(* IEC 61131-3 sources: veristc/veri-stc/tests/st-examples (part 2) *)

cond_a := LimitHigh(raw_030_a, 130);
cond_a := cond_a AND quality_a;
cond_a := cond_a AND (NOT bypass_a);
input_valid_a := InputValid(raw_030_a, 0, 1000);
cond_a := cond_a AND input_valid_a;
IF NOT input_valid_a THEN
    channel_fault_a := channel_fault_a + 1;
END_IF;
cond_b := LimitHigh(raw_030_b, 130);
cond_b := cond_b AND quality_b;
cond_b := cond_b AND (NOT bypass_b);
input_valid_b := InputValid(raw_030_b, 0, 1000);
cond_b := cond_b AND input_valid_b;
IF NOT input_valid_b THEN
    channel_fault_b := channel_fault_b + 1;
END_IF;
cond_c := LimitHigh(raw_030_c, 130);
cond_c := cond_c AND quality_c;
cond_c := cond_c AND (NOT bypass_c);
input_valid_c := InputValid(raw_030_c, 0, 1000);
cond_c := cond_c AND input_valid_c;
IF NOT input_valid_c THEN
    channel_fault_c := channel_fault_c + 1;
END_IF;
cond_d := LimitHigh(raw_030_d, 130);
cond_d := cond_d AND quality_d;
cond_d := cond_d AND (NOT bypass_d);
input_valid_d := InputValid(raw_030_d, 0, 1000);
cond_d := cond_d AND input_valid_d;
IF NOT input_valid_d THEN
    channel_fault_d := channel_fault_d + 1;
END_IF;
vote_ok := TwoOfFour(cond_a, cond_b, cond_c, cond_d);
IF cond_a <> cond_b THEN
    diagnosis_count := diagnosis_count + 1;
END_IF;
IF cond_c <> cond_d THEN
    diagnosis_count := diagnosis_count + 1;
END_IF;
IF NOT vote_ok THEN
    diagnosis_count := diagnosis_count + 1;
END_IF;
latch_a_030 := RS_Next(vote_ok, train_a_reset, latch_a_030);
IF latch_a_030 AND (NOT train_a_inhibit) THEN
    mask_a_03 := mask_a_03 + 64;
    trip_a := 0 < 1;
    scram_a := 0 < 1;
    breaker_a := 0 > 1;
    mfw_a := 0 < 1;
    alarm_a := 0 < 1;
END_IF;
latch_b_030 := RS_Next(vote_ok, train_b_reset, latch_b_030);
IF latch_b_030 AND (NOT train_b_inhibit) THEN
    mask_b_03 := mask_b_03 + 64;
    trip_b := 0 < 1;
    scram_b := 0 < 1;
    breaker_b := 0 > 1;
    mfw_b := 0 < 1;
    alarm_b := 0 < 1;
END_IF;
IF (raw_030_a > 130) AND (NOT cond_a) THEN
    channel_fault_a := channel_fault_a + 1;
END_IF;
IF (raw_030_b > 130) AND (NOT cond_b) THEN
    channel_fault_b := channel_fault_b + 1;
END_IF;
IF (raw_030_c > 130) AND (NOT cond_c) THEN
    channel_fault_c := channel_fault_c + 1;
END_IF;
IF (raw_030_d > 130) AND (NOT cond_d) THEN
    channel_fault_d := channel_fault_d + 1;
END_IF;
IF vote_ok AND train_a_inhibit THEN
    diagnosis_count := diagnosis_count + 1;
END_IF;
IF vote_ok AND train_b_inhibit THEN
    diagnosis_count := diagnosis_count + 1;
END_IF;

cond_a := LimitHigh(raw_031_a, 131);
cond_a := cond_a AND quality_a;
cond_a := cond_a AND (NOT bypass_a);
input_valid_a := InputValid(raw_031_a, 0, 1000);
cond_a := cond_a AND input_valid_a;
IF NOT input_valid_a THEN
    channel_fault_a := channel_fault_a + 1;
END_IF;
cond_b := LimitHigh(raw_031_b, 131);
cond_b := cond_b AND quality_b;
cond_b := cond_b AND (NOT bypass_b);
input_valid_b := InputValid(raw_031_b, 0, 1000);
cond_b := cond_b AND input_valid_b;
IF NOT input_valid_b THEN
    channel_fault_b := channel_fault_b + 1;
END_IF;
cond_c := LimitHigh(raw_031_c, 131);
cond_c := cond_c AND quality_c;
cond_c := cond_c AND (NOT bypass_c);
input_valid_c := InputValid(raw_031_c, 0, 1000);
cond_c := cond_c AND input_valid_c;
IF NOT input_valid_c THEN
    channel_fault_c := channel_fault_c + 1;
END_IF;
cond_d := LimitHigh(raw_031_d, 131);
cond_d := cond_d AND quality_d;
cond_d := cond_d AND (NOT bypass_d);
input_valid_d := InputValid(raw_031_d, 0, 1000);
cond_d := cond_d AND input_valid_d;
IF NOT input_valid_d THEN
    channel_fault_d := channel_fault_d + 1;
END_IF;
vote_ok := TwoOfFour(cond_a, cond_b, cond_c, cond_d);
IF cond_a <> cond_b THEN
    diagnosis_count := diagnosis_count + 1;
END_IF;
IF cond_c <> cond_d THEN
    diagnosis_count := diagnosis_count + 1;
END_IF;
IF NOT vote_ok THEN
    diagnosis_count := diagnosis_count + 1;
END_IF;
latch_a_031 := RS_Next(vote_ok, train_a_reset, latch_a_031);
IF latch_a_031 AND (NOT train_a_inhibit) THEN
    mask_a_03 := mask_a_03 + 128;
    trip_a := 0 < 1;
    scram_a := 0 < 1;
    breaker_a := 0 > 1;
    afw_a := 0 < 1;
    alarm_a := 0 < 1;
END_IF;
latch_b_031 := RS_Next(vote_ok, train_b_reset, latch_b_031);
IF latch_b_031 AND (NOT train_b_inhibit) THEN
    mask_b_03 := mask_b_03 + 128;
    trip_b := 0 < 1;
    scram_b := 0 < 1;
    breaker_b := 0 > 1;
    afw_b := 0 < 1;
    alarm_b := 0 < 1;
END_IF;
IF (raw_031_a > 131) AND (NOT cond_a) THEN
    channel_fault_a := channel_fault_a + 1;
END_IF;
IF (raw_031_b > 131) AND (NOT cond_b) THEN
    channel_fault_b := channel_fault_b + 1;
END_IF;
IF (raw_031_c > 131) AND (NOT cond_c) THEN
    channel_fault_c := channel_fault_c + 1;
END_IF;
IF (raw_031_d > 131) AND (NOT cond_d) THEN
    channel_fault_d := channel_fault_d + 1;
END_IF;
IF vote_ok AND train_a_inhibit THEN
    diagnosis_count := diagnosis_count + 1;
END_IF;
IF vote_ok AND train_b_inhibit THEN
    diagnosis_count := diagnosis_count + 1;
END_IF;

cond_a := LimitHigh(raw_032_a, 132);
cond_a := cond_a AND quality_a;
cond_a := cond_a AND (NOT bypass_a);
input_valid_a := InputValid(raw_032_a, 0, 1000);
cond_a := cond_a AND input_valid_a;
IF NOT input_valid_a THEN
    channel_fault_a := channel_fault_a + 1;
END_IF;
cond_b := LimitHigh(raw_032_b, 132);
cond_b := cond_b AND quality_b;
cond_b := cond_b AND (NOT bypass_b);
input_valid_b := InputValid(raw_032_b, 0, 1000);
cond_b := cond_b AND input_valid_b;
IF NOT input_valid_b THEN
    channel_fault_b := channel_fault_b + 1;
END_IF;
cond_c := LimitHigh(raw_032_c, 132);
cond_c := cond_c AND quality_c;
cond_c := cond_c AND (NOT bypass_c);
input_valid_c := InputValid(raw_032_c, 0, 1000);
cond_c := cond_c AND input_valid_c;
IF NOT input_valid_c THEN
    channel_fault_c := channel_fault_c + 1;
END_IF;
cond_d := LimitHigh(raw_032_d, 132);
cond_d := cond_d AND quality_d;
cond_d := cond_d AND (NOT bypass_d);
input_valid_d := InputValid(raw_032_d, 0, 1000);
cond_d := cond_d AND input_valid_d;
IF NOT input_valid_d THEN
    channel_fault_d := channel_fault_d + 1;
END_IF;
vote_ok := TwoOfFour(cond_a, cond_b, cond_c, cond_d);
IF cond_a <> cond_b THEN
    diagnosis_count := diagnosis_count + 1;
END_IF;
IF cond_c <> cond_d THEN
    diagnosis_count := diagnosis_count + 1;
END_IF;
IF NOT vote_ok THEN
    diagnosis_count := diagnosis_count + 1;
END_IF;
latch_a_032 := RS_Next(vote_ok, train_a_reset, latch_a_032);
IF latch_a_032 AND (NOT train_a_inhibit) THEN
    mask_a_04 := mask_a_04 + 1;
    trip_a := 0 < 1;
    scram_a := 0 < 1;
    breaker_a := 0 > 1;
    si_a := 0 < 1;
    alarm_a := 0 < 1;
END_IF;
latch_b_032 := RS_Next(vote_ok, train_b_reset, latch_b_032);
IF latch_b_032 AND (NOT train_b_inhibit) THEN
    mask_b_04 := mask_b_04 + 1;
    trip_b := 0 < 1;
    scram_b := 0 < 1;
    breaker_b := 0 > 1;
    si_b := 0 < 1;
    alarm_b := 0 < 1;
END_IF;
IF (raw_032_a > 132) AND (NOT cond_a) THEN
    channel_fault_a := channel_fault_a + 1;
END_IF;
IF (raw_032_b > 132) AND (NOT cond_b) THEN
    channel_fault_b := channel_fault_b + 1;
END_IF;
IF (raw_032_c > 132) AND (NOT cond_c) THEN
    channel_fault_c := channel_fault_c + 1;
END_IF;
IF (raw_032_d > 132) AND (NOT cond_d) THEN
    channel_fault_d := channel_fault_d + 1;
END_IF;
IF vote_ok AND train_a_inhibit THEN
    diagnosis_count := diagnosis_count + 1;
END_IF;
IF vote_ok AND train_b_inhibit THEN
    diagnosis_count := diagnosis_count + 1;
END_IF;

cond_a := LimitHigh(raw_033_a, 133);
cond_a := cond_a AND quality_a;
cond_a := cond_a AND (NOT bypass_a);
input_valid_a := InputValid(raw_033_a, 0, 1000);
cond_a := cond_a AND input_valid_a;
IF NOT input_valid_a THEN
    channel_fault_a := channel_fault_a + 1;
END_IF;
cond_b := LimitHigh(raw_033_b, 133);
cond_b := cond_b AND quality_b;
cond_b := cond_b AND (NOT bypass_b);
input_valid_b := InputValid(raw_033_b, 0, 1000);
cond_b := cond_b AND input_valid_b;
IF NOT input_valid_b THEN
    channel_fault_b := channel_fault_b + 1;
END_IF;
cond_c := LimitHigh(raw_033_c, 133);
cond_c := cond_c AND quality_c;
cond_c := cond_c AND (NOT bypass_c);
input_valid_c := InputValid(raw_033_c, 0, 1000);
cond_c := cond_c AND input_valid_c;
IF NOT input_valid_c THEN
    channel_fault_c := channel_fault_c + 1;
END_IF;
cond_d := LimitHigh(raw_033_d, 133);
cond_d := cond_d AND quality_d;
cond_d := cond_d AND (NOT bypass_d);
input_valid_d := InputValid(raw_033_d, 0, 1000);
cond_d := cond_d AND input_valid_d;
IF NOT input_valid_d THEN
    channel_fault_d := channel_fault_d + 1;
END_IF;
vote_ok := TwoOfFour(cond_a, cond_b, cond_c, cond_d);
IF cond_a <> cond_b THEN
    diagnosis_count := diagnosis_count + 1;
END_IF;
IF cond_c <> cond_d THEN
    diagnosis_count := diagnosis_count + 1;
END_IF;
IF NOT vote_ok THEN
    diagnosis_count := diagnosis_count + 1;
END_IF;
latch_a_033 := RS_Next(vote_ok, train_a_reset, latch_a_033);
IF latch_a_033 AND (NOT train_a_inhibit) THEN
    mask_a_04 := mask_a_04 + 2;
    trip_a := 0 < 1;
    scram_a := 0 < 1;
    breaker_a := 0 > 1;
    ci_a := 0 < 1;
    alarm_a := 0 < 1;
END_IF;
latch_b_033 := RS_Next(vote_ok, train_b_reset, latch_b_033);
IF latch_b_033 AND (NOT train_b_inhibit) THEN
    mask_b_04 := mask_b_04 + 2;
    trip_b := 0 < 1;
    scram_b := 0 < 1;
    breaker_b := 0 > 1;
    ci_b := 0 < 1;
    alarm_b := 0 < 1;
END_IF;
IF (raw_033_a > 133) AND (NOT cond_a) THEN
    channel_fault_a := channel_fault_a + 1;
END_IF;
IF (raw_033_b > 133) AND (NOT cond_b) THEN
    channel_fault_b := channel_fault_b + 1;
END_IF;
IF (raw_033_c > 133) AND (NOT cond_c) THEN
    channel_fault_c := channel_fault_c + 1;
END_IF;
IF (raw_033_d > 133) AND (NOT cond_d) THEN
    channel_fault_d := channel_fault_d + 1;
END_IF;
IF vote_ok AND train_a_inhibit THEN
    diagnosis_count := diagnosis_count + 1;
END_IF;
IF vote_ok AND train_b_inhibit THEN
    diagnosis_count := diagnosis_count + 1;
END_IF;

cond_a := LimitHigh(raw_034_a, 134);
cond_a := cond_a AND quality_a;
cond_a := cond_a AND (NOT bypass_a);
input_valid_a := InputValid(raw_034_a, 0, 1000);
cond_a := cond_a AND input_valid_a;
IF NOT input_valid_a THEN
    channel_fault_a := channel_fault_a + 1;
END_IF;
cond_b := LimitHigh(raw_034_b, 134);
cond_b := cond_b AND quality_b;
cond_b := cond_b AND (NOT bypass_b);
input_valid_b := InputValid(raw_034_b, 0, 1000);
cond_b := cond_b AND input_valid_b;
IF NOT input_valid_b THEN
    channel_fault_b := channel_fault_b + 1;
END_IF;
cond_c := LimitHigh(raw_034_c, 134);
cond_c := cond_c AND quality_c;
cond_c := cond_c AND (NOT bypass_c);
input_valid_c := InputValid(raw_034_c, 0, 1000);
cond_c := cond_c AND input_valid_c;
IF NOT input_valid_c THEN
    channel_fault_c := channel_fault_c + 1;
END_IF;
cond_d := LimitHigh(raw_034_d, 134);
cond_d := cond_d AND quality_d;
cond_d := cond_d AND (NOT bypass_d);
input_valid_d := InputValid(raw_034_d, 0, 1000);
cond_d := cond_d AND input_valid_d;
IF NOT input_valid_d THEN
    channel_fault_d := channel_fault_d + 1;
END_IF;
vote_ok := TwoOfFour(cond_a, cond_b, cond_c, cond_d);
IF cond_a <> cond_b THEN
    diagnosis_count := diagnosis_count + 1;
END_IF;
IF cond_c <> cond_d THEN
    diagnosis_count := diagnosis_count + 1;
END_IF;
IF NOT vote_ok THEN
    diagnosis_count := diagnosis_count + 1;
END_IF;
latch_a_034 := RS_Next(vote_ok, train_a_reset, latch_a_034);
IF latch_a_034 AND (NOT train_a_inhibit) THEN
    mask_a_04 := mask_a_04 + 4;
    trip_a := 0 < 1;
    scram_a := 0 < 1;
    breaker_a := 0 > 1;
    mfw_a := 0 < 1;
    alarm_a := 0 < 1;
END_IF;
latch_b_034 := RS_Next(vote_ok, train_b_reset, latch_b_034);
IF latch_b_034 AND (NOT train_b_inhibit) THEN
    mask_b_04 := mask_b_04 + 4;
    trip_b := 0 < 1;
    scram_b := 0 < 1;
    breaker_b := 0 > 1;
    mfw_b := 0 < 1;
    alarm_b := 0 < 1;
END_IF;
IF (raw_034_a > 134) AND (NOT cond_a) THEN
    channel_fault_a := channel_fault_a + 1;
END_IF;
IF (raw_034_b > 134) AND (NOT cond_b) THEN
    channel_fault_b := channel_fault_b + 1;
END_IF;
IF (raw_034_c > 134) AND (NOT cond_c) THEN
    channel_fault_c := channel_fault_c + 1;
END_IF;
IF (raw_034_d > 134) AND (NOT cond_d) THEN
    channel_fault_d := channel_fault_d + 1;
END_IF;
IF vote_ok AND train_a_inhibit THEN
    diagnosis_count := diagnosis_count + 1;
END_IF;
IF vote_ok AND train_b_inhibit THEN
    diagnosis_count := diagnosis_count + 1;
END_IF;

cond_a := LimitHigh(raw_035_a, 135);
cond_a := cond_a AND quality_a;
cond_a := cond_a AND (NOT bypass_a);
input_valid_a := InputValid(raw_035_a, 0, 1000);
cond_a := cond_a AND input_valid_a;
IF NOT input_valid_a THEN
    channel_fault_a := channel_fault_a + 1;
END_IF;
cond_b := LimitHigh(raw_035_b, 135);
cond_b := cond_b AND quality_b;
cond_b := cond_b AND (NOT bypass_b);
input_valid_b := InputValid(raw_035_b, 0, 1000);
cond_b := cond_b AND input_valid_b;
IF NOT input_valid_b THEN
    channel_fault_b := channel_fault_b + 1;
END_IF;
cond_c := LimitHigh(raw_035_c, 135);
cond_c := cond_c AND quality_c;
cond_c := cond_c AND (NOT bypass_c);
input_valid_c := InputValid(raw_035_c, 0, 1000);
cond_c := cond_c AND input_valid_c;
IF NOT input_valid_c THEN
    channel_fault_c := channel_fault_c + 1;
END_IF;
cond_d := LimitHigh(raw_035_d, 135);
cond_d := cond_d AND quality_d;
cond_d := cond_d AND (NOT bypass_d);
input_valid_d := InputValid(raw_035_d, 0, 1000);
cond_d := cond_d AND input_valid_d;
IF NOT input_valid_d THEN
    channel_fault_d := channel_fault_d + 1;
END_IF;
vote_ok := TwoOfFour(cond_a, cond_b, cond_c, cond_d);
IF cond_a <> cond_b THEN
    diagnosis_count := diagnosis_count + 1;
END_IF;
IF cond_c <> cond_d THEN
    diagnosis_count := diagnosis_count + 1;
END_IF;
IF NOT vote_ok THEN
    diagnosis_count := diagnosis_count + 1;
END_IF;
latch_a_035 := RS_Next(vote_ok, train_a_reset, latch_a_035);
IF latch_a_035 AND (NOT train_a_inhibit) THEN
    mask_a_04 := mask_a_04 + 8;
    trip_a := 0 < 1;
    scram_a := 0 < 1;
    breaker_a := 0 > 1;
    afw_a := 0 < 1;
    alarm_a := 0 < 1;
END_IF;
latch_b_035 := RS_Next(vote_ok, train_b_reset, latch_b_035);
IF latch_b_035 AND (NOT train_b_inhibit) THEN
    mask_b_04 := mask_b_04 + 8;
    trip_b := 0 < 1;
    scram_b := 0 < 1;
    breaker_b := 0 > 1;
    afw_b := 0 < 1;
    alarm_b := 0 < 1;
END_IF;
IF (raw_035_a > 135) AND (NOT cond_a) THEN
    channel_fault_a := channel_fault_a + 1;
END_IF;
IF (raw_035_b > 135) AND (NOT cond_b) THEN
    channel_fault_b := channel_fault_b + 1;
END_IF;
IF (raw_035_c > 135) AND (NOT cond_c) THEN
    channel_fault_c := channel_fault_c + 1;
END_IF;
IF (raw_035_d > 135) AND (NOT cond_d) THEN
    channel_fault_d := channel_fault_d + 1;
END_IF;
IF vote_ok AND train_a_inhibit THEN
    diagnosis_count := diagnosis_count + 1;
END_IF;
IF vote_ok AND train_b_inhibit THEN
    diagnosis_count := diagnosis_count + 1;
END_IF;

cond_a := LimitHigh(raw_036_a, 136);
cond_a := cond_a AND quality_a;
cond_a := cond_a AND (NOT bypass_a);
input_valid_a := InputValid(raw_036_a, 0, 1000);
cond_a := cond_a AND input_valid_a;
IF NOT input_valid_a THEN
    channel_fault_a := channel_fault_a + 1;
END_IF;
cond_b := LimitHigh(raw_036_b, 136);
cond_b := cond_b AND quality_b;
cond_b := cond_b AND (NOT bypass_b);
input_valid_b := InputValid(raw_036_b, 0, 1000);
cond_b := cond_b AND input_valid_b;
IF NOT input_valid_b THEN
    channel_fault_b := channel_fault_b + 1;
END_IF;
cond_c := LimitHigh(raw_036_c, 136);
cond_c := cond_c AND quality_c;
cond_c := cond_c AND (NOT bypass_c);
input_valid_c := InputValid(raw_036_c, 0, 1000);
cond_c := cond_c AND input_valid_c;
IF NOT input_valid_c THEN
    channel_fault_c := channel_fault_c + 1;
END_IF;
cond_d := LimitHigh(raw_036_d, 136);
cond_d := cond_d AND quality_d;
cond_d := cond_d AND (NOT bypass_d);
input_valid_d := InputValid(raw_036_d, 0, 1000);
cond_d := cond_d AND input_valid_d;
IF NOT input_valid_d THEN
    channel_fault_d := channel_fault_d + 1;
END_IF;
vote_ok := TwoOfFour(cond_a, cond_b, cond_c, cond_d);
IF cond_a <> cond_b THEN
    diagnosis_count := diagnosis_count + 1;
END_IF;
IF cond_c <> cond_d THEN
    diagnosis_count := diagnosis_count + 1;
END_IF;
IF NOT vote_ok THEN
    diagnosis_count := diagnosis_count + 1;
END_IF;
latch_a_036 := RS_Next(vote_ok, train_a_reset, latch_a_036);
IF latch_a_036 AND (NOT train_a_inhibit) THEN
    mask_a_04 := mask_a_04 + 16;
    trip_a := 0 < 1;
    scram_a := 0 < 1;
    breaker_a := 0 > 1;
    si_a := 0 < 1;
    alarm_a := 0 < 1;
END_IF;
latch_b_036 := RS_Next(vote_ok, train_b_reset, latch_b_036);
IF latch_b_036 AND (NOT train_b_inhibit) THEN
    mask_b_04 := mask_b_04 + 16;
    trip_b := 0 < 1;
    scram_b := 0 < 1;
    breaker_b := 0 > 1;
    si_b := 0 < 1;
    alarm_b := 0 < 1;
END_IF;
IF (raw_036_a > 136) AND (NOT cond_a) THEN
    channel_fault_a := channel_fault_a + 1;
END_IF;
IF (raw_036_b > 136) AND (NOT cond_b) THEN
    channel_fault_b := channel_fault_b + 1;
END_IF;
IF (raw_036_c > 136) AND (NOT cond_c) THEN
    channel_fault_c := channel_fault_c + 1;
END_IF;
IF (raw_036_d > 136) AND (NOT cond_d) THEN
    channel_fault_d := channel_fault_d + 1;
END_IF;
IF vote_ok AND train_a_inhibit THEN
    diagnosis_count := diagnosis_count + 1;
END_IF;
IF vote_ok AND train_b_inhibit THEN
    diagnosis_count := diagnosis_count + 1;
END_IF;

cond_a := LimitHigh(raw_037_a, 137);
cond_a := cond_a AND quality_a;
cond_a := cond_a AND (NOT bypass_a);
input_valid_a := InputValid(raw_037_a, 0, 1000);
cond_a := cond_a AND input_valid_a;
IF NOT input_valid_a THEN
    channel_fault_a := channel_fault_a + 1;
END_IF;
cond_b := LimitHigh(raw_037_b, 137);
cond_b := cond_b AND quality_b;
cond_b := cond_b AND (NOT bypass_b);
input_valid_b := InputValid(raw_037_b, 0, 1000);
cond_b := cond_b AND input_valid_b;
IF NOT input_valid_b THEN
    channel_fault_b := channel_fault_b + 1;
END_IF;
cond_c := LimitHigh(raw_037_c, 137);
cond_c := cond_c AND quality_c;
cond_c := cond_c AND (NOT bypass_c);
input_valid_c := InputValid(raw_037_c, 0, 1000);
cond_c := cond_c AND input_valid_c;
IF NOT input_valid_c THEN
    channel_fault_c := channel_fault_c + 1;
END_IF;
cond_d := LimitHigh(raw_037_d, 137);
cond_d := cond_d AND quality_d;
cond_d := cond_d AND (NOT bypass_d);
input_valid_d := InputValid(raw_037_d, 0, 1000);
cond_d := cond_d AND input_valid_d;
IF NOT input_valid_d THEN
    channel_fault_d := channel_fault_d + 1;
END_IF;
vote_ok := TwoOfFour(cond_a, cond_b, cond_c, cond_d);
IF cond_a <> cond_b THEN
    diagnosis_count := diagnosis_count + 1;
END_IF;
IF cond_c <> cond_d THEN
    diagnosis_count := diagnosis_count + 1;
END_IF;
IF NOT vote_ok THEN
    diagnosis_count := diagnosis_count + 1;
END_IF;
latch_a_037 := RS_Next(vote_ok, train_a_reset, latch_a_037);
IF latch_a_037 AND (NOT train_a_inhibit) THEN
    mask_a_04 := mask_a_04 + 32;
    trip_a := 0 < 1;
    scram_a := 0 < 1;
    breaker_a := 0 > 1;
    ci_a := 0 < 1;
    alarm_a := 0 < 1;
END_IF;
latch_b_037 := RS_Next(vote_ok, train_b_reset, latch_b_037);
IF latch_b_037 AND (NOT train_b_inhibit) THEN
    mask_b_04 := mask_b_04 + 32;
    trip_b := 0 < 1;
    scram_b := 0 < 1;
    breaker_b := 0 > 1;
    ci_b := 0 < 1;
    alarm_b := 0 < 1;
END_IF;
IF (raw_037_a > 137) AND (NOT cond_a) THEN
    channel_fault_a := channel_fault_a + 1;
END_IF;
IF (raw_037_b > 137) AND (NOT cond_b) THEN
    channel_fault_b := channel_fault_b + 1;
END_IF;
IF (raw_037_c > 137) AND (NOT cond_c) THEN
    channel_fault_c := channel_fault_c + 1;
END_IF;
IF (raw_037_d > 137) AND (NOT cond_d) THEN
    channel_fault_d := channel_fault_d + 1;
END_IF;
IF vote_ok AND train_a_inhibit THEN
    diagnosis_count := diagnosis_count + 1;
END_IF;
IF vote_ok AND train_b_inhibit THEN
    diagnosis_count := diagnosis_count + 1;
END_IF;

cond_a := LimitHigh(raw_038_a, 138);
cond_a := cond_a AND quality_a;
cond_a := cond_a AND (NOT bypass_a);
input_valid_a := InputValid(raw_038_a, 0, 1000);
cond_a := cond_a AND input_valid_a;
IF NOT input_valid_a THEN
    channel_fault_a := channel_fault_a + 1;
END_IF;
cond_b := LimitHigh(raw_038_b, 138);
cond_b := cond_b AND quality_b;
cond_b := cond_b AND (NOT bypass_b);
input_valid_b := InputValid(raw_038_b, 0, 1000);
cond_b := cond_b AND input_valid_b;
IF NOT input_valid_b THEN
    channel_fault_b := channel_fault_b + 1;
END_IF;
cond_c := LimitHigh(raw_038_c, 138);
cond_c := cond_c AND quality_c;
cond_c := cond_c AND (NOT bypass_c);
input_valid_c := InputValid(raw_038_c, 0, 1000);
cond_c := cond_c AND input_valid_c;
IF NOT input_valid_c THEN
    channel_fault_c := channel_fault_c + 1;
END_IF;
cond_d := LimitHigh(raw_038_d, 138);
cond_d := cond_d AND quality_d;
cond_d := cond_d AND (NOT bypass_d);
input_valid_d := InputValid(raw_038_d, 0, 1000);
cond_d := cond_d AND input_valid_d;
IF NOT input_valid_d THEN
    channel_fault_d := channel_fault_d + 1;
END_IF;
vote_ok := TwoOfFour(cond_a, cond_b, cond_c, cond_d);
IF cond_a <> cond_b THEN
    diagnosis_count := diagnosis_count + 1;
END_IF;
IF cond_c <> cond_d THEN
    diagnosis_count := diagnosis_count + 1;
END_IF;
IF NOT vote_ok THEN
    diagnosis_count := diagnosis_count + 1;
END_IF;
latch_a_038 := RS_Next(vote_ok, train_a_reset, latch_a_038);
IF latch_a_038 AND (NOT train_a_inhibit) THEN
    mask_a_04 := mask_a_04 + 64;
    trip_a := 0 < 1;
    scram_a := 0 < 1;
    breaker_a := 0 > 1;
    mfw_a := 0 < 1;
    alarm_a := 0 < 1;
END_IF;
latch_b_038 := RS_Next(vote_ok, train_b_reset, latch_b_038);
IF latch_b_038 AND (NOT train_b_inhibit) THEN
    mask_b_04 := mask_b_04 + 64;
    trip_b := 0 < 1;
    scram_b := 0 < 1;
    breaker_b := 0 > 1;
    mfw_b := 0 < 1;
    alarm_b := 0 < 1;
END_IF;
IF (raw_038_a > 138) AND (NOT cond_a) THEN
    channel_fault_a := channel_fault_a + 1;
END_IF;
IF (raw_038_b > 138) AND (NOT cond_b) THEN
    channel_fault_b := channel_fault_b + 1;
END_IF;
IF (raw_038_c > 138) AND (NOT cond_c) THEN
    channel_fault_c := channel_fault_c + 1;
END_IF;
IF (raw_038_d > 138) AND (NOT cond_d) THEN
    channel_fault_d := channel_fault_d + 1;
END_IF;
IF vote_ok AND train_a_inhibit THEN
    diagnosis_count := diagnosis_count + 1;
END_IF;
IF vote_ok AND train_b_inhibit THEN
    diagnosis_count := diagnosis_count + 1;
END_IF;

cond_a := LimitHigh(raw_039_a, 139);
cond_a := cond_a AND quality_a;
cond_a := cond_a AND (NOT bypass_a);
input_valid_a := InputValid(raw_039_a, 0, 1000);
cond_a := cond_a AND input_valid_a;
IF NOT input_valid_a THEN
    channel_fault_a := channel_fault_a + 1;
END_IF;
cond_b := LimitHigh(raw_039_b, 139);
cond_b := cond_b AND quality_b;
cond_b := cond_b AND (NOT bypass_b);
input_valid_b := InputValid(raw_039_b, 0, 1000);
cond_b := cond_b AND input_valid_b;
IF NOT input_valid_b THEN
    channel_fault_b := channel_fault_b + 1;
END_IF;
cond_c := LimitHigh(raw_039_c, 139);
cond_c := cond_c AND quality_c;
cond_c := cond_c AND (NOT bypass_c);
input_valid_c := InputValid(raw_039_c, 0, 1000);
cond_c := cond_c AND input_valid_c;
IF NOT input_valid_c THEN
    channel_fault_c := channel_fault_c + 1;
END_IF;
cond_d := LimitHigh(raw_039_d, 139);
cond_d := cond_d AND quality_d;
cond_d := cond_d AND (NOT bypass_d);
input_valid_d := InputValid(raw_039_d, 0, 1000);
cond_d := cond_d AND input_valid_d;
IF NOT input_valid_d THEN
    channel_fault_d := channel_fault_d + 1;
END_IF;
vote_ok := TwoOfFour(cond_a, cond_b, cond_c, cond_d);
IF cond_a <> cond_b THEN
    diagnosis_count := diagnosis_count + 1;
END_IF;
IF cond_c <> cond_d THEN
    diagnosis_count := diagnosis_count + 1;
END_IF;
IF NOT vote_ok THEN
    diagnosis_count := diagnosis_count + 1;
END_IF;
latch_a_039 := RS_Next(vote_ok, train_a_reset, latch_a_039);
IF latch_a_039 AND (NOT train_a_inhibit) THEN
    mask_a_04 := mask_a_04 + 128;
    trip_a := 0 < 1;
    scram_a := 0 < 1;
    breaker_a := 0 > 1;
    afw_a := 0 < 1;
    alarm_a := 0 < 1;
END_IF;
latch_b_039 := RS_Next(vote_ok, train_b_reset, latch_b_039);
IF latch_b_039 AND (NOT train_b_inhibit) THEN
    mask_b_04 := mask_b_04 + 128;
    trip_b := 0 < 1;
    scram_b := 0 < 1;
    breaker_b := 0 > 1;
    afw_b := 0 < 1;
    alarm_b := 0 < 1;
END_IF;
IF (raw_039_a > 139) AND (NOT cond_a) THEN
    channel_fault_a := channel_fault_a + 1;
END_IF;
IF (raw_039_b > 139) AND (NOT cond_b) THEN
    channel_fault_b := channel_fault_b + 1;
END_IF;
IF (raw_039_c > 139) AND (NOT cond_c) THEN
    channel_fault_c := channel_fault_c + 1;
END_IF;
IF (raw_039_d > 139) AND (NOT cond_d) THEN
    channel_fault_d := channel_fault_d + 1;
END_IF;
IF vote_ok AND train_a_inhibit THEN
    diagnosis_count := diagnosis_count + 1;
END_IF;
IF vote_ok AND train_b_inhibit THEN
    diagnosis_count := diagnosis_count + 1;
END_IF;

cond_a := LimitHigh(raw_040_a, 100);
cond_a := cond_a AND quality_a;
cond_a := cond_a AND (NOT bypass_a);
input_valid_a := InputValid(raw_040_a, 0, 1000);
cond_a := cond_a AND input_valid_a;
IF NOT input_valid_a THEN
    channel_fault_a := channel_fault_a + 1;
END_IF;
cond_b := LimitHigh(raw_040_b, 100);
cond_b := cond_b AND quality_b;
cond_b := cond_b AND (NOT bypass_b);
input_valid_b := InputValid(raw_040_b, 0, 1000);
cond_b := cond_b AND input_valid_b;
IF NOT input_valid_b THEN
    channel_fault_b := channel_fault_b + 1;
END_IF;
cond_c := LimitHigh(raw_040_c, 100);
cond_c := cond_c AND quality_c;
cond_c := cond_c AND (NOT bypass_c);
input_valid_c := InputValid(raw_040_c, 0, 1000);
cond_c := cond_c AND input_valid_c;
IF NOT input_valid_c THEN
    channel_fault_c := channel_fault_c + 1;
END_IF;
cond_d := LimitHigh(raw_040_d, 100);
cond_d := cond_d AND quality_d;
cond_d := cond_d AND (NOT bypass_d);
input_valid_d := InputValid(raw_040_d, 0, 1000);
cond_d := cond_d AND input_valid_d;
IF NOT input_valid_d THEN
    channel_fault_d := channel_fault_d + 1;
END_IF;
vote_ok := TwoOfFour(cond_a, cond_b, cond_c, cond_d);
IF cond_a <> cond_b THEN
    diagnosis_count := diagnosis_count + 1;
END_IF;
IF cond_c <> cond_d THEN
    diagnosis_count := diagnosis_count + 1;
END_IF;
IF NOT vote_ok THEN
    diagnosis_count := diagnosis_count + 1;
END_IF;
latch_a_040 := RS_Next(vote_ok, train_a_reset, latch_a_040);
IF latch_a_040 AND (NOT train_a_inhibit) THEN
    mask_a_05 := mask_a_05 + 1;
    trip_a := 0 < 1;
    scram_a := 0 < 1;
    breaker_a := 0 > 1;
    si_a := 0 < 1;
    alarm_a := 0 < 1;
END_IF;
latch_b_040 := RS_Next(vote_ok, train_b_reset, latch_b_040);
IF latch_b_040 AND (NOT train_b_inhibit) THEN
    mask_b_05 := mask_b_05 + 1;
    trip_b := 0 < 1;
    scram_b := 0 < 1;
    breaker_b := 0 > 1;
    si_b := 0 < 1;
    alarm_b := 0 < 1;
END_IF;
IF (raw_040_a > 100) AND (NOT cond_a) THEN
    channel_fault_a := channel_fault_a + 1;
END_IF;
IF (raw_040_b > 100) AND (NOT cond_b) THEN
    channel_fault_b := channel_fault_b + 1;
END_IF;
IF (raw_040_c > 100) AND (NOT cond_c) THEN
    channel_fault_c := channel_fault_c + 1;
END_IF;
IF (raw_040_d > 100) AND (NOT cond_d) THEN
    channel_fault_d := channel_fault_d + 1;
END_IF;
IF vote_ok AND train_a_inhibit THEN
    diagnosis_count := diagnosis_count + 1;
END_IF;
IF vote_ok AND train_b_inhibit THEN
    diagnosis_count := diagnosis_count + 1;
END_IF;

cond_a := LimitHigh(raw_041_a, 101);
cond_a := cond_a AND quality_a;
cond_a := cond_a AND (NOT bypass_a);
input_valid_a := InputValid(raw_041_a, 0, 1000);
cond_a := cond_a AND input_valid_a;
IF NOT input_valid_a THEN
    channel_fault_a := channel_fault_a + 1;
END_IF;
cond_b := LimitHigh(raw_041_b, 101);
cond_b := cond_b AND quality_b;
cond_b := cond_b AND (NOT bypass_b);
input_valid_b := InputValid(raw_041_b, 0, 1000);
cond_b := cond_b AND input_valid_b;
IF NOT input_valid_b THEN
    channel_fault_b := channel_fault_b + 1;
END_IF;
cond_c := LimitHigh(raw_041_c, 101);
cond_c := cond_c AND quality_c;
cond_c := cond_c AND (NOT bypass_c);
input_valid_c := InputValid(raw_041_c, 0, 1000);
cond_c := cond_c AND input_valid_c;
IF NOT input_valid_c THEN
    channel_fault_c := channel_fault_c + 1;
END_IF;
cond_d := LimitHigh(raw_041_d, 101);
cond_d := cond_d AND quality_d;
cond_d := cond_d AND (NOT bypass_d);
input_valid_d := InputValid(raw_041_d, 0, 1000);
cond_d := cond_d AND input_valid_d;
IF NOT input_valid_d THEN
    channel_fault_d := channel_fault_d + 1;
END_IF;
vote_ok := TwoOfFour(cond_a, cond_b, cond_c, cond_d);
IF cond_a <> cond_b THEN
    diagnosis_count := diagnosis_count + 1;
END_IF;
IF cond_c <> cond_d THEN
    diagnosis_count := diagnosis_count + 1;
END_IF;
IF NOT vote_ok THEN
    diagnosis_count := diagnosis_count + 1;
END_IF;
latch_a_041 := RS_Next(vote_ok, train_a_reset, latch_a_041);
IF latch_a_041 AND (NOT train_a_inhibit) THEN
    mask_a_05 := mask_a_05 + 2;
    trip_a := 0 < 1;
    scram_a := 0 < 1;
    breaker_a := 0 > 1;
    ci_a := 0 < 1;
    alarm_a := 0 < 1;
END_IF;
latch_b_041 := RS_Next(vote_ok, train_b_reset, latch_b_041);
IF latch_b_041 AND (NOT train_b_inhibit) THEN
    mask_b_05 := mask_b_05 + 2;
    trip_b := 0 < 1;
    scram_b := 0 < 1;
    breaker_b := 0 > 1;
    ci_b := 0 < 1;
    alarm_b := 0 < 1;
END_IF;
IF (raw_041_a > 101) AND (NOT cond_a) THEN
    channel_fault_a := channel_fault_a + 1;
END_IF;
IF (raw_041_b > 101) AND (NOT cond_b) THEN
    channel_fault_b := channel_fault_b + 1;
END_IF;
IF (raw_041_c > 101) AND (NOT cond_c) THEN
    channel_fault_c := channel_fault_c + 1;
END_IF;
IF (raw_041_d > 101) AND (NOT cond_d) THEN
    channel_fault_d := channel_fault_d + 1;
END_IF;
IF vote_ok AND train_a_inhibit THEN
    diagnosis_count := diagnosis_count + 1;
END_IF;
IF vote_ok AND train_b_inhibit THEN
    diagnosis_count := diagnosis_count + 1;
END_IF;

cond_a := LimitHigh(raw_042_a, 102);
cond_a := cond_a AND quality_a;
cond_a := cond_a AND (NOT bypass_a);
input_valid_a := InputValid(raw_042_a, 0, 1000);
cond_a := cond_a AND input_valid_a;
IF NOT input_valid_a THEN
    channel_fault_a := channel_fault_a + 1;
END_IF;
cond_b := LimitHigh(raw_042_b, 102);
cond_b := cond_b AND quality_b;
cond_b := cond_b AND (NOT bypass_b);
input_valid_b := InputValid(raw_042_b, 0, 1000);
cond_b := cond_b AND input_valid_b;
IF NOT input_valid_b THEN
    channel_fault_b := channel_fault_b + 1;
END_IF;
cond_c := LimitHigh(raw_042_c, 102);
cond_c := cond_c AND quality_c;
cond_c := cond_c AND (NOT bypass_c);
input_valid_c := InputValid(raw_042_c, 0, 1000);
cond_c := cond_c AND input_valid_c;
IF NOT input_valid_c THEN
    channel_fault_c := channel_fault_c + 1;
END_IF;
cond_d := LimitHigh(raw_042_d, 102);
cond_d := cond_d AND quality_d;
cond_d := cond_d AND (NOT bypass_d);
input_valid_d := InputValid(raw_042_d, 0, 1000);
cond_d := cond_d AND input_valid_d;
IF NOT input_valid_d THEN
    channel_fault_d := channel_fault_d + 1;
END_IF;
vote_ok := TwoOfFour(cond_a, cond_b, cond_c, cond_d);
IF cond_a <> cond_b THEN
    diagnosis_count := diagnosis_count + 1;
END_IF;
IF cond_c <> cond_d THEN
    diagnosis_count := diagnosis_count + 1;
END_IF;
IF NOT vote_ok THEN
    diagnosis_count := diagnosis_count + 1;
END_IF;
latch_a_042 := RS_Next(vote_ok, train_a_reset, latch_a_042);
IF latch_a_042 AND (NOT train_a_inhibit) THEN
    mask_a_05 := mask_a_05 + 4;
    trip_a := 0 < 1;
    scram_a := 0 < 1;
    breaker_a := 0 > 1;
    mfw_a := 0 < 1;
    alarm_a := 0 < 1;
END_IF;
latch_b_042 := RS_Next(vote_ok, train_b_reset, latch_b_042);
IF latch_b_042 AND (NOT train_b_inhibit) THEN
    mask_b_05 := mask_b_05 + 4;
    trip_b := 0 < 1;
    scram_b := 0 < 1;
    breaker_b := 0 > 1;
    mfw_b := 0 < 1;
    alarm_b := 0 < 1;
END_IF;
IF (raw_042_a > 102) AND (NOT cond_a) THEN
    channel_fault_a := channel_fault_a + 1;
END_IF;
IF (raw_042_b > 102) AND (NOT cond_b) THEN
    channel_fault_b := channel_fault_b + 1;
END_IF;
IF (raw_042_c > 102) AND (NOT cond_c) THEN
    channel_fault_c := channel_fault_c + 1;
END_IF;
IF (raw_042_d > 102) AND (NOT cond_d) THEN
    channel_fault_d := channel_fault_d + 1;
END_IF;
IF vote_ok AND train_a_inhibit THEN
    diagnosis_count := diagnosis_count + 1;
END_IF;
IF vote_ok AND train_b_inhibit THEN
    diagnosis_count := diagnosis_count + 1;
END_IF;

cond_a := LimitHigh(raw_043_a, 103);
cond_a := cond_a AND quality_a;
cond_a := cond_a AND (NOT bypass_a);
input_valid_a := InputValid(raw_043_a, 0, 1000);
cond_a := cond_a AND input_valid_a;
IF NOT input_valid_a THEN
    channel_fault_a := channel_fault_a + 1;
END_IF;
cond_b := LimitHigh(raw_043_b, 103);
cond_b := cond_b AND quality_b;
cond_b := cond_b AND (NOT bypass_b);
input_valid_b := InputValid(raw_043_b, 0, 1000);
cond_b := cond_b AND input_valid_b;
IF NOT input_valid_b THEN
    channel_fault_b := channel_fault_b + 1;
END_IF;
cond_c := LimitHigh(raw_043_c, 103);
cond_c := cond_c AND quality_c;
cond_c := cond_c AND (NOT bypass_c);
input_valid_c := InputValid(raw_043_c, 0, 1000);
cond_c := cond_c AND input_valid_c;
IF NOT input_valid_c THEN
    channel_fault_c := channel_fault_c + 1;
END_IF;
cond_d := LimitHigh(raw_043_d, 103);
cond_d := cond_d AND quality_d;
cond_d := cond_d AND (NOT bypass_d);
input_valid_d := InputValid(raw_043_d, 0, 1000);
cond_d := cond_d AND input_valid_d;
IF NOT input_valid_d THEN
    channel_fault_d := channel_fault_d + 1;
END_IF;
vote_ok := TwoOfFour(cond_a, cond_b, cond_c, cond_d);
IF cond_a <> cond_b THEN
    diagnosis_count := diagnosis_count + 1;
END_IF;
IF cond_c <> cond_d THEN
    diagnosis_count := diagnosis_count + 1;
END_IF;
IF NOT vote_ok THEN
    diagnosis_count := diagnosis_count + 1;
END_IF;
latch_a_043 := RS_Next(vote_ok, train_a_reset, latch_a_043);
IF latch_a_043 AND (NOT train_a_inhibit) THEN
    mask_a_05 := mask_a_05 + 8;
    trip_a := 0 < 1;
    scram_a := 0 < 1;
    breaker_a := 0 > 1;
    afw_a := 0 < 1;
    alarm_a := 0 < 1;
END_IF;
latch_b_043 := RS_Next(vote_ok, train_b_reset, latch_b_043);
IF latch_b_043 AND (NOT train_b_inhibit) THEN
    mask_b_05 := mask_b_05 + 8;
    trip_b := 0 < 1;
    scram_b := 0 < 1;
    breaker_b := 0 > 1;
    afw_b := 0 < 1;
    alarm_b := 0 < 1;
END_IF;
IF (raw_043_a > 103) AND (NOT cond_a) THEN
    channel_fault_a := channel_fault_a + 1;
END_IF;
IF (raw_043_b > 103) AND (NOT cond_b) THEN
    channel_fault_b := channel_fault_b + 1;
END_IF;
IF (raw_043_c > 103) AND (NOT cond_c) THEN
    channel_fault_c := channel_fault_c + 1;
END_IF;
IF (raw_043_d > 103) AND (NOT cond_d) THEN
    channel_fault_d := channel_fault_d + 1;
END_IF;
IF vote_ok AND train_a_inhibit THEN
    diagnosis_count := diagnosis_count + 1;
END_IF;
IF vote_ok AND train_b_inhibit THEN
    diagnosis_count := diagnosis_count + 1;
END_IF;

cond_a := LimitHigh(raw_044_a, 104);
cond_a := cond_a AND quality_a;
cond_a := cond_a AND (NOT bypass_a);
input_valid_a := InputValid(raw_044_a, 0, 1000);
cond_a := cond_a AND input_valid_a;
IF NOT input_valid_a THEN
    channel_fault_a := channel_fault_a + 1;
END_IF;
cond_b := LimitHigh(raw_044_b, 104);
cond_b := cond_b AND quality_b;
cond_b := cond_b AND (NOT bypass_b);
input_valid_b := InputValid(raw_044_b, 0, 1000);
cond_b := cond_b AND input_valid_b;
IF NOT input_valid_b THEN
    channel_fault_b := channel_fault_b + 1;
END_IF;
cond_c := LimitHigh(raw_044_c, 104);
cond_c := cond_c AND quality_c;
cond_c := cond_c AND (NOT bypass_c);
input_valid_c := InputValid(raw_044_c, 0, 1000);
cond_c := cond_c AND input_valid_c;
IF NOT input_valid_c THEN
    channel_fault_c := channel_fault_c + 1;
END_IF;
cond_d := LimitHigh(raw_044_d, 104);
cond_d := cond_d AND quality_d;
cond_d := cond_d AND (NOT bypass_d);
input_valid_d := InputValid(raw_044_d, 0, 1000);
cond_d := cond_d AND input_valid_d;
IF NOT input_valid_d THEN
    channel_fault_d := channel_fault_d + 1;
END_IF;
vote_ok := TwoOfFour(cond_a, cond_b, cond_c, cond_d);
IF cond_a <> cond_b THEN
    diagnosis_count := diagnosis_count + 1;
END_IF;
IF cond_c <> cond_d THEN
    diagnosis_count := diagnosis_count + 1;
END_IF;
IF NOT vote_ok THEN
    diagnosis_count := diagnosis_count + 1;
END_IF;
latch_a_044 := RS_Next(vote_ok, train_a_reset, latch_a_044);
IF latch_a_044 AND (NOT train_a_inhibit) THEN
    mask_a_05 := mask_a_05 + 16;
    trip_a := 0 < 1;
    scram_a := 0 < 1;
    breaker_a := 0 > 1;
    si_a := 0 < 1;
    alarm_a := 0 < 1;
END_IF;
latch_b_044 := RS_Next(vote_ok, train_b_reset, latch_b_044);
IF latch_b_044 AND (NOT train_b_inhibit) THEN
    mask_b_05 := mask_b_05 + 16;
    trip_b := 0 < 1;
    scram_b := 0 < 1;
    breaker_b := 0 > 1;
    si_b := 0 < 1;
    alarm_b := 0 < 1;
END_IF;
IF (raw_044_a > 104) AND (NOT cond_a) THEN
    channel_fault_a := channel_fault_a + 1;
END_IF;
IF (raw_044_b > 104) AND (NOT cond_b) THEN
    channel_fault_b := channel_fault_b + 1;
END_IF;
IF (raw_044_c > 104) AND (NOT cond_c) THEN
    channel_fault_c := channel_fault_c + 1;
END_IF;
IF (raw_044_d > 104) AND (NOT cond_d) THEN
    channel_fault_d := channel_fault_d + 1;
END_IF;
IF vote_ok AND train_a_inhibit THEN
    diagnosis_count := diagnosis_count + 1;
END_IF;
IF vote_ok AND train_b_inhibit THEN
    diagnosis_count := diagnosis_count + 1;
END_IF;

cond_a := LimitHigh(raw_045_a, 105);
cond_a := cond_a AND quality_a;
cond_a := cond_a AND (NOT bypass_a);
input_valid_a := InputValid(raw_045_a, 0, 1000);
cond_a := cond_a AND input_valid_a;
IF NOT input_valid_a THEN
    channel_fault_a := channel_fault_a + 1;
END_IF;
cond_b := LimitHigh(raw_045_b, 105);
cond_b := cond_b AND quality_b;
cond_b := cond_b AND (NOT bypass_b);
input_valid_b := InputValid(raw_045_b, 0, 1000);
cond_b := cond_b AND input_valid_b;
IF NOT input_valid_b THEN
    channel_fault_b := channel_fault_b + 1;
END_IF;
cond_c := LimitHigh(raw_045_c, 105);
cond_c := cond_c AND quality_c;
cond_c := cond_c AND (NOT bypass_c);
input_valid_c := InputValid(raw_045_c, 0, 1000);
cond_c := cond_c AND input_valid_c;
IF NOT input_valid_c THEN
    channel_fault_c := channel_fault_c + 1;
END_IF;
cond_d := LimitHigh(raw_045_d, 105);
cond_d := cond_d AND quality_d;
cond_d := cond_d AND (NOT bypass_d);
input_valid_d := InputValid(raw_045_d, 0, 1000);
cond_d := cond_d AND input_valid_d;
IF NOT input_valid_d THEN
    channel_fault_d := channel_fault_d + 1;
END_IF;
vote_ok := TwoOfFour(cond_a, cond_b, cond_c, cond_d);
IF cond_a <> cond_b THEN
    diagnosis_count := diagnosis_count + 1;
END_IF;
IF cond_c <> cond_d THEN
    diagnosis_count := diagnosis_count + 1;
END_IF;
IF NOT vote_ok THEN
    diagnosis_count := diagnosis_count + 1;
END_IF;
latch_a_045 := RS_Next(vote_ok, train_a_reset, latch_a_045);
IF latch_a_045 AND (NOT train_a_inhibit) THEN
    mask_a_05 := mask_a_05 + 32;
    trip_a := 0 < 1;
    scram_a := 0 < 1;
    breaker_a := 0 > 1;
    ci_a := 0 < 1;
    alarm_a := 0 < 1;
END_IF;
latch_b_045 := RS_Next(vote_ok, train_b_reset, latch_b_045);
IF latch_b_045 AND (NOT train_b_inhibit) THEN
    mask_b_05 := mask_b_05 + 32;
    trip_b := 0 < 1;
    scram_b := 0 < 1;
    breaker_b := 0 > 1;
    ci_b := 0 < 1;
    alarm_b := 0 < 1;
END_IF;
IF (raw_045_a > 105) AND (NOT cond_a) THEN
    channel_fault_a := channel_fault_a + 1;
END_IF;
IF (raw_045_b > 105) AND (NOT cond_b) THEN
    channel_fault_b := channel_fault_b + 1;
END_IF;
IF (raw_045_c > 105) AND (NOT cond_c) THEN
    channel_fault_c := channel_fault_c + 1;
END_IF;
IF (raw_045_d > 105) AND (NOT cond_d) THEN
    channel_fault_d := channel_fault_d + 1;
END_IF;
IF vote_ok AND train_a_inhibit THEN
    diagnosis_count := diagnosis_count + 1;
END_IF;
IF vote_ok AND train_b_inhibit THEN
    diagnosis_count := diagnosis_count + 1;
END_IF;

cond_a := LimitHigh(raw_046_a, 106);
cond_a := cond_a AND quality_a;
cond_a := cond_a AND (NOT bypass_a);
input_valid_a := InputValid(raw_046_a, 0, 1000);
cond_a := cond_a AND input_valid_a;
IF NOT input_valid_a THEN
    channel_fault_a := channel_fault_a + 1;
END_IF;
cond_b := LimitHigh(raw_046_b, 106);
cond_b := cond_b AND quality_b;
cond_b := cond_b AND (NOT bypass_b);
input_valid_b := InputValid(raw_046_b, 0, 1000);
cond_b := cond_b AND input_valid_b;
IF NOT input_valid_b THEN
    channel_fault_b := channel_fault_b + 1;
END_IF;
cond_c := LimitHigh(raw_046_c, 106);
cond_c := cond_c AND quality_c;
cond_c := cond_c AND (NOT bypass_c);
input_valid_c := InputValid(raw_046_c, 0, 1000);
cond_c := cond_c AND input_valid_c;
IF NOT input_valid_c THEN
    channel_fault_c := channel_fault_c + 1;
END_IF;
cond_d := LimitHigh(raw_046_d, 106);
cond_d := cond_d AND quality_d;
cond_d := cond_d AND (NOT bypass_d);
input_valid_d := InputValid(raw_046_d, 0, 1000);
cond_d := cond_d AND input_valid_d;
IF NOT input_valid_d THEN
    channel_fault_d := channel_fault_d + 1;
END_IF;
vote_ok := TwoOfFour(cond_a, cond_b, cond_c, cond_d);
IF cond_a <> cond_b THEN
    diagnosis_count := diagnosis_count + 1;
END_IF;
IF cond_c <> cond_d THEN
    diagnosis_count := diagnosis_count + 1;
END_IF;
IF NOT vote_ok THEN
    diagnosis_count := diagnosis_count + 1;
END_IF;
latch_a_046 := RS_Next(vote_ok, train_a_reset, latch_a_046);
IF latch_a_046 AND (NOT train_a_inhibit) THEN
    mask_a_05 := mask_a_05 + 64;
    trip_a := 0 < 1;
    scram_a := 0 < 1;
    breaker_a := 0 > 1;
    mfw_a := 0 < 1;
    alarm_a := 0 < 1;
END_IF;
latch_b_046 := RS_Next(vote_ok, train_b_reset, latch_b_046);
IF latch_b_046 AND (NOT train_b_inhibit) THEN
    mask_b_05 := mask_b_05 + 64;
    trip_b := 0 < 1;
    scram_b := 0 < 1;
    breaker_b := 0 > 1;
    mfw_b := 0 < 1;
    alarm_b := 0 < 1;
END_IF;
IF (raw_046_a > 106) AND (NOT cond_a) THEN
    channel_fault_a := channel_fault_a + 1;
END_IF;
IF (raw_046_b > 106) AND (NOT cond_b) THEN
    channel_fault_b := channel_fault_b + 1;
END_IF;
IF (raw_046_c > 106) AND (NOT cond_c) THEN
    channel_fault_c := channel_fault_c + 1;
END_IF;
IF (raw_046_d > 106) AND (NOT cond_d) THEN
    channel_fault_d := channel_fault_d + 1;
END_IF;
IF vote_ok AND train_a_inhibit THEN
    diagnosis_count := diagnosis_count + 1;
END_IF;
IF vote_ok AND train_b_inhibit THEN
    diagnosis_count := diagnosis_count + 1;
END_IF;

cond_a := LimitHigh(raw_047_a, 107);
cond_a := cond_a AND quality_a;
cond_a := cond_a AND (NOT bypass_a);
input_valid_a := InputValid(raw_047_a, 0, 1000);
cond_a := cond_a AND input_valid_a;
IF NOT input_valid_a THEN
    channel_fault_a := channel_fault_a + 1;
END_IF;
cond_b := LimitHigh(raw_047_b, 107);
cond_b := cond_b AND quality_b;
cond_b := cond_b AND (NOT bypass_b);
input_valid_b := InputValid(raw_047_b, 0, 1000);
cond_b := cond_b AND input_valid_b;
IF NOT input_valid_b THEN
    channel_fault_b := channel_fault_b + 1;
END_IF;
cond_c := LimitHigh(raw_047_c, 107);
cond_c := cond_c AND quality_c;
cond_c := cond_c AND (NOT bypass_c);
input_valid_c := InputValid(raw_047_c, 0, 1000);
cond_c := cond_c AND input_valid_c;
IF NOT input_valid_c THEN
    channel_fault_c := channel_fault_c + 1;
END_IF;
cond_d := LimitHigh(raw_047_d, 107);
cond_d := cond_d AND quality_d;
cond_d := cond_d AND (NOT bypass_d);
input_valid_d := InputValid(raw_047_d, 0, 1000);
cond_d := cond_d AND input_valid_d;
IF NOT input_valid_d THEN
    channel_fault_d := channel_fault_d + 1;
END_IF;
vote_ok := TwoOfFour(cond_a, cond_b, cond_c, cond_d);
IF cond_a <> cond_b THEN
    diagnosis_count := diagnosis_count + 1;
END_IF;
IF cond_c <> cond_d THEN
    diagnosis_count := diagnosis_count + 1;
END_IF;
IF NOT vote_ok THEN
    diagnosis_count := diagnosis_count + 1;
END_IF;
latch_a_047 := RS_Next(vote_ok, train_a_reset, latch_a_047);
IF latch_a_047 AND (NOT train_a_inhibit) THEN
    mask_a_05 := mask_a_05 + 128;
    trip_a := 0 < 1;
    scram_a := 0 < 1;
    breaker_a := 0 > 1;
    afw_a := 0 < 1;
    alarm_a := 0 < 1;
END_IF;
latch_b_047 := RS_Next(vote_ok, train_b_reset, latch_b_047);
IF latch_b_047 AND (NOT train_b_inhibit) THEN
    mask_b_05 := mask_b_05 + 128;
    trip_b := 0 < 1;
    scram_b := 0 < 1;
    breaker_b := 0 > 1;
    afw_b := 0 < 1;
    alarm_b := 0 < 1;
END_IF;
IF (raw_047_a > 107) AND (NOT cond_a) THEN
    channel_fault_a := channel_fault_a + 1;
END_IF;
IF (raw_047_b > 107) AND (NOT cond_b) THEN
    channel_fault_b := channel_fault_b + 1;
END_IF;
IF (raw_047_c > 107) AND (NOT cond_c) THEN
    channel_fault_c := channel_fault_c + 1;
END_IF;
IF (raw_047_d > 107) AND (NOT cond_d) THEN
    channel_fault_d := channel_fault_d + 1;
END_IF;
IF vote_ok AND train_a_inhibit THEN
    diagnosis_count := diagnosis_count + 1;
END_IF;
IF vote_ok AND train_b_inhibit THEN
    diagnosis_count := diagnosis_count + 1;
END_IF;

cond_a := LimitHigh(raw_048_a, 108);
cond_a := cond_a AND quality_a;
cond_a := cond_a AND (NOT bypass_a);
input_valid_a := InputValid(raw_048_a, 0, 1000);
cond_a := cond_a AND input_valid_a;
IF NOT input_valid_a THEN
    channel_fault_a := channel_fault_a + 1;
END_IF;
cond_b := LimitHigh(raw_048_b, 108);
cond_b := cond_b AND quality_b;
cond_b := cond_b AND (NOT bypass_b);
input_valid_b := InputValid(raw_048_b, 0, 1000);
cond_b := cond_b AND input_valid_b;
IF NOT input_valid_b THEN
    channel_fault_b := channel_fault_b + 1;
END_IF;
cond_c := LimitHigh(raw_048_c, 108);
cond_c := cond_c AND quality_c;
cond_c := cond_c AND (NOT bypass_c);
input_valid_c := InputValid(raw_048_c, 0, 1000);
cond_c := cond_c AND input_valid_c;
IF NOT input_valid_c THEN
    channel_fault_c := channel_fault_c + 1;
END_IF;
cond_d := LimitHigh(raw_048_d, 108);
cond_d := cond_d AND quality_d;
cond_d := cond_d AND (NOT bypass_d);
input_valid_d := InputValid(raw_048_d, 0, 1000);
cond_d := cond_d AND input_valid_d;
IF NOT input_valid_d THEN
    channel_fault_d := channel_fault_d + 1;
END_IF;
vote_ok := TwoOfFour(cond_a, cond_b, cond_c, cond_d);
IF cond_a <> cond_b THEN
    diagnosis_count := diagnosis_count + 1;
END_IF;
IF cond_c <> cond_d THEN
    diagnosis_count := diagnosis_count + 1;
END_IF;
IF NOT vote_ok THEN
    diagnosis_count := diagnosis_count + 1;
END_IF;
latch_a_048 := RS_Next(vote_ok, train_a_reset, latch_a_048);
IF latch_a_048 AND (NOT train_a_inhibit) THEN
    mask_a_06 := mask_a_06 + 1;
    trip_a := 0 < 1;
    scram_a := 0 < 1;
    breaker_a := 0 > 1;
    si_a := 0 < 1;
    alarm_a := 0 < 1;
END_IF;
latch_b_048 := RS_Next(vote_ok, train_b_reset, latch_b_048);
IF latch_b_048 AND (NOT train_b_inhibit) THEN
    mask_b_06 := mask_b_06 + 1;
    trip_b := 0 < 1;
    scram_b := 0 < 1;
    breaker_b := 0 > 1;
    si_b := 0 < 1;
    alarm_b := 0 < 1;
END_IF;
IF (raw_048_a > 108) AND (NOT cond_a) THEN
    channel_fault_a := channel_fault_a + 1;
END_IF;
IF (raw_048_b > 108) AND (NOT cond_b) THEN
    channel_fault_b := channel_fault_b + 1;
END_IF;
IF (raw_048_c > 108) AND (NOT cond_c) THEN
    channel_fault_c := channel_fault_c + 1;
END_IF;
IF (raw_048_d > 108) AND (NOT cond_d) THEN
    channel_fault_d := channel_fault_d + 1;
END_IF;
IF vote_ok AND train_a_inhibit THEN
    diagnosis_count := diagnosis_count + 1;
END_IF;
IF vote_ok AND train_b_inhibit THEN
    diagnosis_count := diagnosis_count + 1;
END_IF;

cond_a := LimitHigh(raw_049_a, 109);
cond_a := cond_a AND quality_a;
cond_a := cond_a AND (NOT bypass_a);
input_valid_a := InputValid(raw_049_a, 0, 1000);
cond_a := cond_a AND input_valid_a;
IF NOT input_valid_a THEN
    channel_fault_a := channel_fault_a + 1;
END_IF;
cond_b := LimitHigh(raw_049_b, 109);
cond_b := cond_b AND quality_b;
cond_b := cond_b AND (NOT bypass_b);
input_valid_b := InputValid(raw_049_b, 0, 1000);
cond_b := cond_b AND input_valid_b;
IF NOT input_valid_b THEN
    channel_fault_b := channel_fault_b + 1;
END_IF;
cond_c := LimitHigh(raw_049_c, 109);
cond_c := cond_c AND quality_c;
cond_c := cond_c AND (NOT bypass_c);
input_valid_c := InputValid(raw_049_c, 0, 1000);
cond_c := cond_c AND input_valid_c;
IF NOT input_valid_c THEN
    channel_fault_c := channel_fault_c + 1;
END_IF;
cond_d := LimitHigh(raw_049_d, 109);
cond_d := cond_d AND quality_d;
cond_d := cond_d AND (NOT bypass_d);
input_valid_d := InputValid(raw_049_d, 0, 1000);
cond_d := cond_d AND input_valid_d;
IF NOT input_valid_d THEN
    channel_fault_d := channel_fault_d + 1;
END_IF;
vote_ok := TwoOfFour(cond_a, cond_b, cond_c, cond_d);
IF cond_a <> cond_b THEN
    diagnosis_count := diagnosis_count + 1;
END_IF;
IF cond_c <> cond_d THEN
    diagnosis_count := diagnosis_count + 1;
END_IF;
IF NOT vote_ok THEN
    diagnosis_count := diagnosis_count + 1;
END_IF;
latch_a_049 := RS_Next(vote_ok, train_a_reset, latch_a_049);
IF latch_a_049 AND (NOT train_a_inhibit) THEN
    mask_a_06 := mask_a_06 + 2;
    trip_a := 0 < 1;
    scram_a := 0 < 1;
    breaker_a := 0 > 1;
    ci_a := 0 < 1;
    alarm_a := 0 < 1;
END_IF;
latch_b_049 := RS_Next(vote_ok, train_b_reset, latch_b_049);
IF latch_b_049 AND (NOT train_b_inhibit) THEN
    mask_b_06 := mask_b_06 + 2;
    trip_b := 0 < 1;
    scram_b := 0 < 1;
    breaker_b := 0 > 1;
    ci_b := 0 < 1;
    alarm_b := 0 < 1;
END_IF;
IF (raw_049_a > 109) AND (NOT cond_a) THEN
    channel_fault_a := channel_fault_a + 1;
END_IF;
IF (raw_049_b > 109) AND (NOT cond_b) THEN
    channel_fault_b := channel_fault_b + 1;
END_IF;
IF (raw_049_c > 109) AND (NOT cond_c) THEN
    channel_fault_c := channel_fault_c + 1;
END_IF;
IF (raw_049_d > 109) AND (NOT cond_d) THEN
    channel_fault_d := channel_fault_d + 1;
END_IF;
IF vote_ok AND train_a_inhibit THEN
    diagnosis_count := diagnosis_count + 1;
END_IF;
IF vote_ok AND train_b_inhibit THEN
    diagnosis_count := diagnosis_count + 1;
END_IF;

cond_a := LimitHigh(raw_050_a, 110);
cond_a := cond_a AND quality_a;
cond_a := cond_a AND (NOT bypass_a);
input_valid_a := InputValid(raw_050_a, 0, 1000);
cond_a := cond_a AND input_valid_a;
IF NOT input_valid_a THEN
    channel_fault_a := channel_fault_a + 1;
END_IF;
cond_b := LimitHigh(raw_050_b, 110);
cond_b := cond_b AND quality_b;
cond_b := cond_b AND (NOT bypass_b);
input_valid_b := InputValid(raw_050_b, 0, 1000);
cond_b := cond_b AND input_valid_b;
IF NOT input_valid_b THEN
    channel_fault_b := channel_fault_b + 1;
END_IF;
cond_c := LimitHigh(raw_050_c, 110);
cond_c := cond_c AND quality_c;
cond_c := cond_c AND (NOT bypass_c);
input_valid_c := InputValid(raw_050_c, 0, 1000);
cond_c := cond_c AND input_valid_c;
IF NOT input_valid_c THEN
    channel_fault_c := channel_fault_c + 1;
END_IF;
cond_d := LimitHigh(raw_050_d, 110);
cond_d := cond_d AND quality_d;
cond_d := cond_d AND (NOT bypass_d);
input_valid_d := InputValid(raw_050_d, 0, 1000);
cond_d := cond_d AND input_valid_d;
IF NOT input_valid_d THEN
    channel_fault_d := channel_fault_d + 1;
END_IF;
vote_ok := TwoOfFour(cond_a, cond_b, cond_c, cond_d);
IF cond_a <> cond_b THEN
    diagnosis_count := diagnosis_count + 1;
END_IF;
IF cond_c <> cond_d THEN
    diagnosis_count := diagnosis_count + 1;
END_IF;
IF NOT vote_ok THEN
    diagnosis_count := diagnosis_count + 1;
END_IF;
latch_a_050 := RS_Next(vote_ok, train_a_reset, latch_a_050);
IF latch_a_050 AND (NOT train_a_inhibit) THEN
    mask_a_06 := mask_a_06 + 4;
    trip_a := 0 < 1;
    scram_a := 0 < 1;
    breaker_a := 0 > 1;
    mfw_a := 0 < 1;
    alarm_a := 0 < 1;
END_IF;
latch_b_050 := RS_Next(vote_ok, train_b_reset, latch_b_050);
IF latch_b_050 AND (NOT train_b_inhibit) THEN
    mask_b_06 := mask_b_06 + 4;
    trip_b := 0 < 1;
    scram_b := 0 < 1;
    breaker_b := 0 > 1;
    mfw_b := 0 < 1;
    alarm_b := 0 < 1;
END_IF;
IF (raw_050_a > 110) AND (NOT cond_a) THEN
    channel_fault_a := channel_fault_a + 1;
END_IF;
IF (raw_050_b > 110) AND (NOT cond_b) THEN
    channel_fault_b := channel_fault_b + 1;
END_IF;
IF (raw_050_c > 110) AND (NOT cond_c) THEN
    channel_fault_c := channel_fault_c + 1;
END_IF;
IF (raw_050_d > 110) AND (NOT cond_d) THEN
    channel_fault_d := channel_fault_d + 1;
END_IF;
IF vote_ok AND train_a_inhibit THEN
    diagnosis_count := diagnosis_count + 1;
END_IF;
IF vote_ok AND train_b_inhibit THEN
    diagnosis_count := diagnosis_count + 1;
END_IF;

cond_a := LimitHigh(raw_051_a, 111);
cond_a := cond_a AND quality_a;
cond_a := cond_a AND (NOT bypass_a);
input_valid_a := InputValid(raw_051_a, 0, 1000);
cond_a := cond_a AND input_valid_a;
IF NOT input_valid_a THEN
    channel_fault_a := channel_fault_a + 1;
END_IF;
cond_b := LimitHigh(raw_051_b, 111);
cond_b := cond_b AND quality_b;
cond_b := cond_b AND (NOT bypass_b);
input_valid_b := InputValid(raw_051_b, 0, 1000);
cond_b := cond_b AND input_valid_b;
IF NOT input_valid_b THEN
    channel_fault_b := channel_fault_b + 1;
END_IF;
cond_c := LimitHigh(raw_051_c, 111);
cond_c := cond_c AND quality_c;
cond_c := cond_c AND (NOT bypass_c);
input_valid_c := InputValid(raw_051_c, 0, 1000);
cond_c := cond_c AND input_valid_c;
IF NOT input_valid_c THEN
    channel_fault_c := channel_fault_c + 1;
END_IF;
cond_d := LimitHigh(raw_051_d, 111);
cond_d := cond_d AND quality_d;
cond_d := cond_d AND (NOT bypass_d);
input_valid_d := InputValid(raw_051_d, 0, 1000);
cond_d := cond_d AND input_valid_d;
IF NOT input_valid_d THEN
    channel_fault_d := channel_fault_d + 1;
END_IF;
vote_ok := TwoOfFour(cond_a, cond_b, cond_c, cond_d);
IF cond_a <> cond_b THEN
    diagnosis_count := diagnosis_count + 1;
END_IF;
IF cond_c <> cond_d THEN
    diagnosis_count := diagnosis_count + 1;
END_IF;
IF NOT vote_ok THEN
    diagnosis_count := diagnosis_count + 1;
END_IF;
latch_a_051 := RS_Next(vote_ok, train_a_reset, latch_a_051);
IF latch_a_051 AND (NOT train_a_inhibit) THEN
    mask_a_06 := mask_a_06 + 8;
    trip_a := 0 < 1;
    scram_a := 0 < 1;
    breaker_a := 0 > 1;
    afw_a := 0 < 1;
    alarm_a := 0 < 1;
END_IF;
latch_b_051 := RS_Next(vote_ok, train_b_reset, latch_b_051);
IF latch_b_051 AND (NOT train_b_inhibit) THEN
    mask_b_06 := mask_b_06 + 8;
    trip_b := 0 < 1;
    scram_b := 0 < 1;
    breaker_b := 0 > 1;
    afw_b := 0 < 1;
    alarm_b := 0 < 1;
END_IF;
IF (raw_051_a > 111) AND (NOT cond_a) THEN
    channel_fault_a := channel_fault_a + 1;
END_IF;
IF (raw_051_b > 111) AND (NOT cond_b) THEN
    channel_fault_b := channel_fault_b + 1;
END_IF;
IF (raw_051_c > 111) AND (NOT cond_c) THEN
    channel_fault_c := channel_fault_c + 1;
END_IF;
IF (raw_051_d > 111) AND (NOT cond_d) THEN
    channel_fault_d := channel_fault_d + 1;
END_IF;
IF vote_ok AND train_a_inhibit THEN
    diagnosis_count := diagnosis_count + 1;
END_IF;
IF vote_ok AND train_b_inhibit THEN
    diagnosis_count := diagnosis_count + 1;
END_IF;

cond_a := LimitHigh(raw_052_a, 112);
cond_a := cond_a AND quality_a;
cond_a := cond_a AND (NOT bypass_a);
input_valid_a := InputValid(raw_052_a, 0, 1000);
cond_a := cond_a AND input_valid_a;
IF NOT input_valid_a THEN
    channel_fault_a := channel_fault_a + 1;
END_IF;
cond_b := LimitHigh(raw_052_b, 112);
cond_b := cond_b AND quality_b;
cond_b := cond_b AND (NOT bypass_b);
input_valid_b := InputValid(raw_052_b, 0, 1000);
cond_b := cond_b AND input_valid_b;
IF NOT input_valid_b THEN
    channel_fault_b := channel_fault_b + 1;
END_IF;
cond_c := LimitHigh(raw_052_c, 112);
cond_c := cond_c AND quality_c;
cond_c := cond_c AND (NOT bypass_c);
input_valid_c := InputValid(raw_052_c, 0, 1000);
cond_c := cond_c AND input_valid_c;
IF NOT input_valid_c THEN
    channel_fault_c := channel_fault_c + 1;
END_IF;
cond_d := LimitHigh(raw_052_d, 112);
cond_d := cond_d AND quality_d;
cond_d := cond_d AND (NOT bypass_d);
input_valid_d := InputValid(raw_052_d, 0, 1000);
cond_d := cond_d AND input_valid_d;
IF NOT input_valid_d THEN
    channel_fault_d := channel_fault_d + 1;
END_IF;
vote_ok := TwoOfFour(cond_a, cond_b, cond_c, cond_d);
IF cond_a <> cond_b THEN
    diagnosis_count := diagnosis_count + 1;
END_IF;
IF cond_c <> cond_d THEN
    diagnosis_count := diagnosis_count + 1;
END_IF;
IF NOT vote_ok THEN
    diagnosis_count := diagnosis_count + 1;
END_IF;
latch_a_052 := RS_Next(vote_ok, train_a_reset, latch_a_052);
IF latch_a_052 AND (NOT train_a_inhibit) THEN
    mask_a_06 := mask_a_06 + 16;
    trip_a := 0 < 1;
    scram_a := 0 < 1;
    breaker_a := 0 > 1;
    si_a := 0 < 1;
    alarm_a := 0 < 1;
END_IF;
latch_b_052 := RS_Next(vote_ok, train_b_reset, latch_b_052);
IF latch_b_052 AND (NOT train_b_inhibit) THEN
    mask_b_06 := mask_b_06 + 16;
    trip_b := 0 < 1;
    scram_b := 0 < 1;
    breaker_b := 0 > 1;
    si_b := 0 < 1;
    alarm_b := 0 < 1;
END_IF;
IF (raw_052_a > 112) AND (NOT cond_a) THEN
    channel_fault_a := channel_fault_a + 1;
END_IF;
IF (raw_052_b > 112) AND (NOT cond_b) THEN
    channel_fault_b := channel_fault_b + 1;
END_IF;
IF (raw_052_c > 112) AND (NOT cond_c) THEN
    channel_fault_c := channel_fault_c + 1;
END_IF;
IF (raw_052_d > 112) AND (NOT cond_d) THEN
    channel_fault_d := channel_fault_d + 1;
END_IF;
IF vote_ok AND train_a_inhibit THEN
    diagnosis_count := diagnosis_count + 1;
END_IF;
IF vote_ok AND train_b_inhibit THEN
    diagnosis_count := diagnosis_count + 1;
END_IF;

cond_a := LimitHigh(raw_053_a, 113);
cond_a := cond_a AND quality_a;
cond_a := cond_a AND (NOT bypass_a);
input_valid_a := InputValid(raw_053_a, 0, 1000);
cond_a := cond_a AND input_valid_a;
IF NOT input_valid_a THEN
    channel_fault_a := channel_fault_a + 1;
END_IF;
cond_b := LimitHigh(raw_053_b, 113);
cond_b := cond_b AND quality_b;
cond_b := cond_b AND (NOT bypass_b);
input_valid_b := InputValid(raw_053_b, 0, 1000);
cond_b := cond_b AND input_valid_b;
IF NOT input_valid_b THEN
    channel_fault_b := channel_fault_b + 1;
END_IF;
cond_c := LimitHigh(raw_053_c, 113);
cond_c := cond_c AND quality_c;
cond_c := cond_c AND (NOT bypass_c);
input_valid_c := InputValid(raw_053_c, 0, 1000);
cond_c := cond_c AND input_valid_c;
IF NOT input_valid_c THEN
    channel_fault_c := channel_fault_c + 1;
END_IF;
cond_d := LimitHigh(raw_053_d, 113);
cond_d := cond_d AND quality_d;
cond_d := cond_d AND (NOT bypass_d);
input_valid_d := InputValid(raw_053_d, 0, 1000);
cond_d := cond_d AND input_valid_d;
IF NOT input_valid_d THEN
    channel_fault_d := channel_fault_d + 1;
END_IF;
vote_ok := TwoOfFour(cond_a, cond_b, cond_c, cond_d);
IF cond_a <> cond_b THEN
    diagnosis_count := diagnosis_count + 1;
END_IF;
IF cond_c <> cond_d THEN
    diagnosis_count := diagnosis_count + 1;
END_IF;
IF NOT vote_ok THEN
    diagnosis_count := diagnosis_count + 1;
END_IF;
latch_a_053 := RS_Next(vote_ok, train_a_reset, latch_a_053);
IF latch_a_053 AND (NOT train_a_inhibit) THEN
    mask_a_06 := mask_a_06 + 32;
    trip_a := 0 < 1;
    scram_a := 0 < 1;
    breaker_a := 0 > 1;
    ci_a := 0 < 1;
    alarm_a := 0 < 1;
END_IF;
latch_b_053 := RS_Next(vote_ok, train_b_reset, latch_b_053);
IF latch_b_053 AND (NOT train_b_inhibit) THEN
    mask_b_06 := mask_b_06 + 32;
    trip_b := 0 < 1;
    scram_b := 0 < 1;
    breaker_b := 0 > 1;
    ci_b := 0 < 1;
    alarm_b := 0 < 1;
END_IF;
IF (raw_053_a > 113) AND (NOT cond_a) THEN
    channel_fault_a := channel_fault_a + 1;
END_IF;
IF (raw_053_b > 113) AND (NOT cond_b) THEN
    channel_fault_b := channel_fault_b + 1;
END_IF;
IF (raw_053_c > 113) AND (NOT cond_c) THEN
    channel_fault_c := channel_fault_c + 1;
END_IF;
IF (raw_053_d > 113) AND (NOT cond_d) THEN
    channel_fault_d := channel_fault_d + 1;
END_IF;
IF vote_ok AND train_a_inhibit THEN
    diagnosis_count := diagnosis_count + 1;
END_IF;
IF vote_ok AND train_b_inhibit THEN
    diagnosis_count := diagnosis_count + 1;
END_IF;

cond_a := LimitHigh(raw_054_a, 114);
cond_a := cond_a AND quality_a;
cond_a := cond_a AND (NOT bypass_a);
input_valid_a := InputValid(raw_054_a, 0, 1000);
cond_a := cond_a AND input_valid_a;
IF NOT input_valid_a THEN
    channel_fault_a := channel_fault_a + 1;
END_IF;
cond_b := LimitHigh(raw_054_b, 114);
cond_b := cond_b AND quality_b;
cond_b := cond_b AND (NOT bypass_b);
input_valid_b := InputValid(raw_054_b, 0, 1000);
cond_b := cond_b AND input_valid_b;
IF NOT input_valid_b THEN
    channel_fault_b := channel_fault_b + 1;
END_IF;
cond_c := LimitHigh(raw_054_c, 114);
cond_c := cond_c AND quality_c;
cond_c := cond_c AND (NOT bypass_c);
input_valid_c := InputValid(raw_054_c, 0, 1000);
cond_c := cond_c AND input_valid_c;
IF NOT input_valid_c THEN
    channel_fault_c := channel_fault_c + 1;
END_IF;
cond_d := LimitHigh(raw_054_d, 114);
cond_d := cond_d AND quality_d;
cond_d := cond_d AND (NOT bypass_d);
input_valid_d := InputValid(raw_054_d, 0, 1000);
cond_d := cond_d AND input_valid_d;
IF NOT input_valid_d THEN
    channel_fault_d := channel_fault_d + 1;
END_IF;
vote_ok := TwoOfFour(cond_a, cond_b, cond_c, cond_d);
IF cond_a <> cond_b THEN
    diagnosis_count := diagnosis_count + 1;
END_IF;
IF cond_c <> cond_d THEN
    diagnosis_count := diagnosis_count + 1;
END_IF;
IF NOT vote_ok THEN
    diagnosis_count := diagnosis_count + 1;
END_IF;
latch_a_054 := RS_Next(vote_ok, train_a_reset, latch_a_054);
IF latch_a_054 AND (NOT train_a_inhibit) THEN
    mask_a_06 := mask_a_06 + 64;
    trip_a := 0 < 1;
    scram_a := 0 < 1;
    breaker_a := 0 > 1;
    mfw_a := 0 < 1;
    alarm_a := 0 < 1;
END_IF;
latch_b_054 := RS_Next(vote_ok, train_b_reset, latch_b_054);
IF latch_b_054 AND (NOT train_b_inhibit) THEN
    mask_b_06 := mask_b_06 + 64;
    trip_b := 0 < 1;
    scram_b := 0 < 1;
    breaker_b := 0 > 1;
    mfw_b := 0 < 1;
    alarm_b := 0 < 1;
END_IF;
IF (raw_054_a > 114) AND (NOT cond_a) THEN
    channel_fault_a := channel_fault_a + 1;
END_IF;
IF (raw_054_b > 114) AND (NOT cond_b) THEN
    channel_fault_b := channel_fault_b + 1;
END_IF;
IF (raw_054_c > 114) AND (NOT cond_c) THEN
    channel_fault_c := channel_fault_c + 1;
END_IF;
IF (raw_054_d > 114) AND (NOT cond_d) THEN
    channel_fault_d := channel_fault_d + 1;
END_IF;
IF vote_ok AND train_a_inhibit THEN
    diagnosis_count := diagnosis_count + 1;
END_IF;
IF vote_ok AND train_b_inhibit THEN
    diagnosis_count := diagnosis_count + 1;
END_IF;

cond_a := LimitHigh(raw_055_a, 115);
cond_a := cond_a AND quality_a;
cond_a := cond_a AND (NOT bypass_a);
input_valid_a := InputValid(raw_055_a, 0, 1000);
cond_a := cond_a AND input_valid_a;
IF NOT input_valid_a THEN
    channel_fault_a := channel_fault_a + 1;
END_IF;
cond_b := LimitHigh(raw_055_b, 115);
cond_b := cond_b AND quality_b;
cond_b := cond_b AND (NOT bypass_b);
input_valid_b := InputValid(raw_055_b, 0, 1000);
cond_b := cond_b AND input_valid_b;
IF NOT input_valid_b THEN
    channel_fault_b := channel_fault_b + 1;
END_IF;
cond_c := LimitHigh(raw_055_c, 115);
cond_c := cond_c AND quality_c;
cond_c := cond_c AND (NOT bypass_c);
input_valid_c := InputValid(raw_055_c, 0, 1000);
cond_c := cond_c AND input_valid_c;
IF NOT input_valid_c THEN
    channel_fault_c := channel_fault_c + 1;
END_IF;
cond_d := LimitHigh(raw_055_d, 115);
cond_d := cond_d AND quality_d;
cond_d := cond_d AND (NOT bypass_d);
input_valid_d := InputValid(raw_055_d, 0, 1000);
cond_d := cond_d AND input_valid_d;
IF NOT input_valid_d THEN
    channel_fault_d := channel_fault_d + 1;
END_IF;
vote_ok := TwoOfFour(cond_a, cond_b, cond_c, cond_d);
IF cond_a <> cond_b THEN
    diagnosis_count := diagnosis_count + 1;
END_IF;
IF cond_c <> cond_d THEN
    diagnosis_count := diagnosis_count + 1;
END_IF;
IF NOT vote_ok THEN
    diagnosis_count := diagnosis_count + 1;
END_IF;
latch_a_055 := RS_Next(vote_ok, train_a_reset, latch_a_055);
IF latch_a_055 AND (NOT train_a_inhibit) THEN
    mask_a_06 := mask_a_06 + 128;
    trip_a := 0 < 1;
    scram_a := 0 < 1;
    breaker_a := 0 > 1;
    afw_a := 0 < 1;
    alarm_a := 0 < 1;
END_IF;
latch_b_055 := RS_Next(vote_ok, train_b_reset, latch_b_055);
IF latch_b_055 AND (NOT train_b_inhibit) THEN
    mask_b_06 := mask_b_06 + 128;
    trip_b := 0 < 1;
    scram_b := 0 < 1;
    breaker_b := 0 > 1;
    afw_b := 0 < 1;
    alarm_b := 0 < 1;
END_IF;
IF (raw_055_a > 115) AND (NOT cond_a) THEN
    channel_fault_a := channel_fault_a + 1;
END_IF;
IF (raw_055_b > 115) AND (NOT cond_b) THEN
    channel_fault_b := channel_fault_b + 1;
END_IF;
IF (raw_055_c > 115) AND (NOT cond_c) THEN
    channel_fault_c := channel_fault_c + 1;
END_IF;
IF (raw_055_d > 115) AND (NOT cond_d) THEN
    channel_fault_d := channel_fault_d + 1;
END_IF;
IF vote_ok AND train_a_inhibit THEN
    diagnosis_count := diagnosis_count + 1;
END_IF;
IF vote_ok AND train_b_inhibit THEN
    diagnosis_count := diagnosis_count + 1;
END_IF;

cond_a := LimitHigh(raw_056_a, 116);
cond_a := cond_a AND quality_a;
cond_a := cond_a AND (NOT bypass_a);
input_valid_a := InputValid(raw_056_a, 0, 1000);
cond_a := cond_a AND input_valid_a;
IF NOT input_valid_a THEN
    channel_fault_a := channel_fault_a + 1;
END_IF;
cond_b := LimitHigh(raw_056_b, 116);
cond_b := cond_b AND quality_b;
cond_b := cond_b AND (NOT bypass_b);
input_valid_b := InputValid(raw_056_b, 0, 1000);
cond_b := cond_b AND input_valid_b;
IF NOT input_valid_b THEN
    channel_fault_b := channel_fault_b + 1;
END_IF;
cond_c := LimitHigh(raw_056_c, 116);
cond_c := cond_c AND quality_c;
cond_c := cond_c AND (NOT bypass_c);
input_valid_c := InputValid(raw_056_c, 0, 1000);
cond_c := cond_c AND input_valid_c;
IF NOT input_valid_c THEN
    channel_fault_c := channel_fault_c + 1;
END_IF;
cond_d := LimitHigh(raw_056_d, 116);
cond_d := cond_d AND quality_d;
cond_d := cond_d AND (NOT bypass_d);
input_valid_d := InputValid(raw_056_d, 0, 1000);
cond_d := cond_d AND input_valid_d;
IF NOT input_valid_d THEN
    channel_fault_d := channel_fault_d + 1;
END_IF;
vote_ok := TwoOfFour(cond_a, cond_b, cond_c, cond_d);
IF cond_a <> cond_b THEN
    diagnosis_count := diagnosis_count + 1;
END_IF;
IF cond_c <> cond_d THEN
    diagnosis_count := diagnosis_count + 1;
END_IF;
IF NOT vote_ok THEN
    diagnosis_count := diagnosis_count + 1;
END_IF;
latch_a_056 := RS_Next(vote_ok, train_a_reset, latch_a_056);
IF latch_a_056 AND (NOT train_a_inhibit) THEN
    mask_a_07 := mask_a_07 + 1;
    trip_a := 0 < 1;
    scram_a := 0 < 1;
    breaker_a := 0 > 1;
    si_a := 0 < 1;
    alarm_a := 0 < 1;
END_IF;
latch_b_056 := RS_Next(vote_ok, train_b_reset, latch_b_056);
IF latch_b_056 AND (NOT train_b_inhibit) THEN
    mask_b_07 := mask_b_07 + 1;
    trip_b := 0 < 1;
    scram_b := 0 < 1;
    breaker_b := 0 > 1;
    si_b := 0 < 1;
    alarm_b := 0 < 1;
END_IF;
IF (raw_056_a > 116) AND (NOT cond_a) THEN
    channel_fault_a := channel_fault_a + 1;
END_IF;
IF (raw_056_b > 116) AND (NOT cond_b) THEN
    channel_fault_b := channel_fault_b + 1;
END_IF;
IF (raw_056_c > 116) AND (NOT cond_c) THEN
    channel_fault_c := channel_fault_c + 1;
END_IF;
IF (raw_056_d > 116) AND (NOT cond_d) THEN
    channel_fault_d := channel_fault_d + 1;
END_IF;
IF vote_ok AND train_a_inhibit THEN
    diagnosis_count := diagnosis_count + 1;
END_IF;
IF vote_ok AND train_b_inhibit THEN
    diagnosis_count := diagnosis_count + 1;
END_IF;

cond_a := LimitHigh(raw_057_a, 117);
cond_a := cond_a AND quality_a;
cond_a := cond_a AND (NOT bypass_a);
input_valid_a := InputValid(raw_057_a, 0, 1000);
cond_a := cond_a AND input_valid_a;
IF NOT input_valid_a THEN
    channel_fault_a := channel_fault_a + 1;
END_IF;
cond_b := LimitHigh(raw_057_b, 117);
cond_b := cond_b AND quality_b;
cond_b := cond_b AND (NOT bypass_b);
input_valid_b := InputValid(raw_057_b, 0, 1000);
cond_b := cond_b AND input_valid_b;
IF NOT input_valid_b THEN
    channel_fault_b := channel_fault_b + 1;
END_IF;
cond_c := LimitHigh(raw_057_c, 117);
cond_c := cond_c AND quality_c;
cond_c := cond_c AND (NOT bypass_c);
input_valid_c := InputValid(raw_057_c, 0, 1000);
cond_c := cond_c AND input_valid_c;
IF NOT input_valid_c THEN
    channel_fault_c := channel_fault_c + 1;
END_IF;
cond_d := LimitHigh(raw_057_d, 117);
cond_d := cond_d AND quality_d;
cond_d := cond_d AND (NOT bypass_d);
input_valid_d := InputValid(raw_057_d, 0, 1000);
cond_d := cond_d AND input_valid_d;
IF NOT input_valid_d THEN
    channel_fault_d := channel_fault_d + 1;
END_IF;
vote_ok := TwoOfFour(cond_a, cond_b, cond_c, cond_d);
IF cond_a <> cond_b THEN
    diagnosis_count := diagnosis_count + 1;
END_IF;
IF cond_c <> cond_d THEN
    diagnosis_count := diagnosis_count + 1;
END_IF;
IF NOT vote_ok THEN
    diagnosis_count := diagnosis_count + 1;
END_IF;
latch_a_057 := RS_Next(vote_ok, train_a_reset, latch_a_057);
IF latch_a_057 AND (NOT train_a_inhibit) THEN
    mask_a_07 := mask_a_07 + 2;
    trip_a := 0 < 1;
    scram_a := 0 < 1;
    breaker_a := 0 > 1;
    ci_a := 0 < 1;
    alarm_a := 0 < 1;
END_IF;
latch_b_057 := RS_Next(vote_ok, train_b_reset, latch_b_057);
IF latch_b_057 AND (NOT train_b_inhibit) THEN
    mask_b_07 := mask_b_07 + 2;
    trip_b := 0 < 1;
    scram_b := 0 < 1;
    breaker_b := 0 > 1;
    ci_b := 0 < 1;
    alarm_b := 0 < 1;
END_IF;
IF (raw_057_a > 117) AND (NOT cond_a) THEN
    channel_fault_a := channel_fault_a + 1;
END_IF;
IF (raw_057_b > 117) AND (NOT cond_b) THEN
    channel_fault_b := channel_fault_b + 1;
END_IF;
IF (raw_057_c > 117) AND (NOT cond_c) THEN
    channel_fault_c := channel_fault_c + 1;
END_IF;
IF (raw_057_d > 117) AND (NOT cond_d) THEN
    channel_fault_d := channel_fault_d + 1;
END_IF;
IF vote_ok AND train_a_inhibit THEN
    diagnosis_count := diagnosis_count + 1;
END_IF;
IF vote_ok AND train_b_inhibit THEN
    diagnosis_count := diagnosis_count + 1;
END_IF;

cond_a := LimitHigh(raw_058_a, 118);
cond_a := cond_a AND quality_a;
cond_a := cond_a AND (NOT bypass_a);
input_valid_a := InputValid(raw_058_a, 0, 1000);
cond_a := cond_a AND input_valid_a;
IF NOT input_valid_a THEN
    channel_fault_a := channel_fault_a + 1;
END_IF;
cond_b := LimitHigh(raw_058_b, 118);
cond_b := cond_b AND quality_b;
cond_b := cond_b AND (NOT bypass_b);
input_valid_b := InputValid(raw_058_b, 0, 1000);
cond_b := cond_b AND input_valid_b;
IF NOT input_valid_b THEN
    channel_fault_b := channel_fault_b + 1;
END_IF;
cond_c := LimitHigh(raw_058_c, 118);
cond_c := cond_c AND quality_c;
cond_c := cond_c AND (NOT bypass_c);
input_valid_c := InputValid(raw_058_c, 0, 1000);
cond_c := cond_c AND input_valid_c;
IF NOT input_valid_c THEN
    channel_fault_c := channel_fault_c + 1;
END_IF;
cond_d := LimitHigh(raw_058_d, 118);
cond_d := cond_d AND quality_d;
cond_d := cond_d AND (NOT bypass_d);
input_valid_d := InputValid(raw_058_d, 0, 1000);
cond_d := cond_d AND input_valid_d;
IF NOT input_valid_d THEN
    channel_fault_d := channel_fault_d + 1;
END_IF;
vote_ok := TwoOfFour(cond_a, cond_b, cond_c, cond_d);
IF cond_a <> cond_b THEN
    diagnosis_count := diagnosis_count + 1;
END_IF;
IF cond_c <> cond_d THEN
    diagnosis_count := diagnosis_count + 1;
END_IF;
IF NOT vote_ok THEN
    diagnosis_count := diagnosis_count + 1;
END_IF;
latch_a_058 := RS_Next(vote_ok, train_a_reset, latch_a_058);
IF latch_a_058 AND (NOT train_a_inhibit) THEN
    mask_a_07 := mask_a_07 + 4;
    trip_a := 0 < 1;
    scram_a := 0 < 1;
    breaker_a := 0 > 1;
    mfw_a := 0 < 1;
    alarm_a := 0 < 1;
END_IF;
latch_b_058 := RS_Next(vote_ok, train_b_reset, latch_b_058);
IF latch_b_058 AND (NOT train_b_inhibit) THEN
    mask_b_07 := mask_b_07 + 4;
    trip_b := 0 < 1;
    scram_b := 0 < 1;
    breaker_b := 0 > 1;
    mfw_b := 0 < 1;
    alarm_b := 0 < 1;
END_IF;
IF (raw_058_a > 118) AND (NOT cond_a) THEN
    channel_fault_a := channel_fault_a + 1;
END_IF;
IF (raw_058_b > 118) AND (NOT cond_b) THEN
    channel_fault_b := channel_fault_b + 1;
END_IF;
IF (raw_058_c > 118) AND (NOT cond_c) THEN
    channel_fault_c := channel_fault_c + 1;
END_IF;
IF (raw_058_d > 118) AND (NOT cond_d) THEN
    channel_fault_d := channel_fault_d + 1;
END_IF;
IF vote_ok AND train_a_inhibit THEN
    diagnosis_count := diagnosis_count + 1;
END_IF;
IF vote_ok AND train_b_inhibit THEN
    diagnosis_count := diagnosis_count + 1;
END_IF;

cond_a := LimitHigh(raw_059_a, 119);
cond_a := cond_a AND quality_a;
cond_a := cond_a AND (NOT bypass_a);
input_valid_a := InputValid(raw_059_a, 0, 1000);
cond_a := cond_a AND input_valid_a;
IF NOT input_valid_a THEN
    channel_fault_a := channel_fault_a + 1;
END_IF;
cond_b := LimitHigh(raw_059_b, 119);
cond_b := cond_b AND quality_b;
cond_b := cond_b AND (NOT bypass_b);
input_valid_b := InputValid(raw_059_b, 0, 1000);
cond_b := cond_b AND input_valid_b;
IF NOT input_valid_b THEN
    channel_fault_b := channel_fault_b + 1;
END_IF;
cond_c := LimitHigh(raw_059_c, 119);
cond_c := cond_c AND quality_c;
cond_c := cond_c AND (NOT bypass_c);
input_valid_c := InputValid(raw_059_c, 0, 1000);
cond_c := cond_c AND input_valid_c;
IF NOT input_valid_c THEN
    channel_fault_c := channel_fault_c + 1;
END_IF;
cond_d := LimitHigh(raw_059_d, 119);
cond_d := cond_d AND quality_d;
cond_d := cond_d AND (NOT bypass_d);
input_valid_d := InputValid(raw_059_d, 0, 1000);
cond_d := cond_d AND input_valid_d;
IF NOT input_valid_d THEN
    channel_fault_d := channel_fault_d + 1;
END_IF;
vote_ok := TwoOfFour(cond_a, cond_b, cond_c, cond_d);
IF cond_a <> cond_b THEN
    diagnosis_count := diagnosis_count + 1;
END_IF;
IF cond_c <> cond_d THEN
    diagnosis_count := diagnosis_count + 1;
END_IF;
IF NOT vote_ok THEN
    diagnosis_count := diagnosis_count + 1;
END_IF;
latch_a_059 := RS_Next(vote_ok, train_a_reset, latch_a_059);
IF latch_a_059 AND (NOT train_a_inhibit) THEN
    mask_a_07 := mask_a_07 + 8;
    trip_a := 0 < 1;
    scram_a := 0 < 1;
    breaker_a := 0 > 1;
    afw_a := 0 < 1;
    alarm_a := 0 < 1;
END_IF;
latch_b_059 := RS_Next(vote_ok, train_b_reset, latch_b_059);
IF latch_b_059 AND (NOT train_b_inhibit) THEN
    mask_b_07 := mask_b_07 + 8;
    trip_b := 0 < 1;
    scram_b := 0 < 1;
    breaker_b := 0 > 1;
    afw_b := 0 < 1;
    alarm_b := 0 < 1;
END_IF;
IF (raw_059_a > 119) AND (NOT cond_a) THEN
    channel_fault_a := channel_fault_a + 1;
END_IF;
IF (raw_059_b > 119) AND (NOT cond_b) THEN
    channel_fault_b := channel_fault_b + 1;
END_IF;
IF (raw_059_c > 119) AND (NOT cond_c) THEN
    channel_fault_c := channel_fault_c + 1;
END_IF;
IF (raw_059_d > 119) AND (NOT cond_d) THEN
    channel_fault_d := channel_fault_d + 1;
END_IF;
IF vote_ok AND train_a_inhibit THEN
    diagnosis_count := diagnosis_count + 1;
END_IF;
IF vote_ok AND train_b_inhibit THEN
    diagnosis_count := diagnosis_count + 1;
END_IF;

cond_a := LimitHigh(raw_060_a, 120);
cond_a := cond_a AND quality_a;
cond_a := cond_a AND (NOT bypass_a);
input_valid_a := InputValid(raw_060_a, 0, 1000);
cond_a := cond_a AND input_valid_a;
IF NOT input_valid_a THEN
    channel_fault_a := channel_fault_a + 1;
END_IF;
cond_b := LimitHigh(raw_060_b, 120);
cond_b := cond_b AND quality_b;
cond_b := cond_b AND (NOT bypass_b);
input_valid_b := InputValid(raw_060_b, 0, 1000);
cond_b := cond_b AND input_valid_b;
IF NOT input_valid_b THEN
    channel_fault_b := channel_fault_b + 1;
END_IF;
cond_c := LimitHigh(raw_060_c, 120);
cond_c := cond_c AND quality_c;
cond_c := cond_c AND (NOT bypass_c);
input_valid_c := InputValid(raw_060_c, 0, 1000);
cond_c := cond_c AND input_valid_c;
IF NOT input_valid_c THEN
    channel_fault_c := channel_fault_c + 1;
END_IF;
cond_d := LimitHigh(raw_060_d, 120);
cond_d := cond_d AND quality_d;
cond_d := cond_d AND (NOT bypass_d);
input_valid_d := InputValid(raw_060_d, 0, 1000);
cond_d := cond_d AND input_valid_d;
IF NOT input_valid_d THEN
    channel_fault_d := channel_fault_d + 1;
END_IF;
vote_ok := TwoOfFour(cond_a, cond_b, cond_c, cond_d);
IF cond_a <> cond_b THEN
    diagnosis_count := diagnosis_count + 1;
END_IF;
IF cond_c <> cond_d THEN
    diagnosis_count := diagnosis_count + 1;
END_IF;
IF NOT vote_ok THEN
    diagnosis_count := diagnosis_count + 1;
END_IF;
latch_a_060 := RS_Next(vote_ok, train_a_reset, latch_a_060);
IF latch_a_060 AND (NOT train_a_inhibit) THEN
    mask_a_07 := mask_a_07 + 16;
    trip_a := 0 < 1;
    scram_a := 0 < 1;
    breaker_a := 0 > 1;
    si_a := 0 < 1;
    alarm_a := 0 < 1;
END_IF;
latch_b_060 := RS_Next(vote_ok, train_b_reset, latch_b_060);
IF latch_b_060 AND (NOT train_b_inhibit) THEN
    mask_b_07 := mask_b_07 + 16;
    trip_b := 0 < 1;
    scram_b := 0 < 1;
    breaker_b := 0 > 1;
    si_b := 0 < 1;
    alarm_b := 0 < 1;
END_IF;
IF (raw_060_a > 120) AND (NOT cond_a) THEN
    channel_fault_a := channel_fault_a + 1;
END_IF;
IF (raw_060_b > 120) AND (NOT cond_b) THEN
    channel_fault_b := channel_fault_b + 1;
END_IF;
IF (raw_060_c > 120) AND (NOT cond_c) THEN
    channel_fault_c := channel_fault_c + 1;
END_IF;
IF (raw_060_d > 120) AND (NOT cond_d) THEN
    channel_fault_d := channel_fault_d + 1;
END_IF;
IF vote_ok AND train_a_inhibit THEN
    diagnosis_count := diagnosis_count + 1;
END_IF;
IF vote_ok AND train_b_inhibit THEN
    diagnosis_count := diagnosis_count + 1;
END_IF;

cond_a := LimitHigh(raw_061_a, 121);
cond_a := cond_a AND quality_a;
cond_a := cond_a AND (NOT bypass_a);
input_valid_a := InputValid(raw_061_a, 0, 1000);
cond_a := cond_a AND input_valid_a;
IF NOT input_valid_a THEN
    channel_fault_a := channel_fault_a + 1;
END_IF;
cond_b := LimitHigh(raw_061_b, 121);
cond_b := cond_b AND quality_b;
cond_b := cond_b AND (NOT bypass_b);
input_valid_b := InputValid(raw_061_b, 0, 1000);
cond_b := cond_b AND input_valid_b;
IF NOT input_valid_b THEN
    channel_fault_b := channel_fault_b + 1;
END_IF;
cond_c := LimitHigh(raw_061_c, 121);
cond_c := cond_c AND quality_c;
cond_c := cond_c AND (NOT bypass_c);
input_valid_c := InputValid(raw_061_c, 0, 1000);
cond_c := cond_c AND input_valid_c;
IF NOT input_valid_c THEN
    channel_fault_c := channel_fault_c + 1;
END_IF;
cond_d := LimitHigh(raw_061_d, 121);
cond_d := cond_d AND quality_d;
cond_d := cond_d AND (NOT bypass_d);
input_valid_d := InputValid(raw_061_d, 0, 1000);
cond_d := cond_d AND input_valid_d;
IF NOT input_valid_d THEN
    channel_fault_d := channel_fault_d + 1;
END_IF;
vote_ok := TwoOfFour(cond_a, cond_b, cond_c, cond_d);
IF cond_a <> cond_b THEN
    diagnosis_count := diagnosis_count + 1;
END_IF;
IF cond_c <> cond_d THEN
    diagnosis_count := diagnosis_count + 1;
END_IF;
IF NOT vote_ok THEN
    diagnosis_count := diagnosis_count + 1;
END_IF;
latch_a_061 := RS_Next(vote_ok, train_a_reset, latch_a_061);
IF latch_a_061 AND (NOT train_a_inhibit) THEN
    mask_a_07 := mask_a_07 + 32;
    trip_a := 0 < 1;
    scram_a := 0 < 1;
    breaker_a := 0 > 1;
    ci_a := 0 < 1;
    alarm_a := 0 < 1;
END_IF;
latch_b_061 := RS_Next(vote_ok, train_b_reset, latch_b_061);
IF latch_b_061 AND (NOT train_b_inhibit) THEN
    mask_b_07 := mask_b_07 + 32;
    trip_b := 0 < 1;
    scram_b := 0 < 1;
    breaker_b := 0 > 1;
    ci_b := 0 < 1;
    alarm_b := 0 < 1;
END_IF;
IF (raw_061_a > 121) AND (NOT cond_a) THEN
    channel_fault_a := channel_fault_a + 1;
END_IF;
IF (raw_061_b > 121) AND (NOT cond_b) THEN
    channel_fault_b := channel_fault_b + 1;
END_IF;
IF (raw_061_c > 121) AND (NOT cond_c) THEN
    channel_fault_c := channel_fault_c + 1;
END_IF;
IF (raw_061_d > 121) AND (NOT cond_d) THEN
    channel_fault_d := channel_fault_d + 1;
END_IF;
IF vote_ok AND train_a_inhibit THEN
    diagnosis_count := diagnosis_count + 1;
END_IF;
IF vote_ok AND train_b_inhibit THEN
    diagnosis_count := diagnosis_count + 1;
END_IF;

cond_a := LimitHigh(raw_062_a, 122);
cond_a := cond_a AND quality_a;
cond_a := cond_a AND (NOT bypass_a);
input_valid_a := InputValid(raw_062_a, 0, 1000);
cond_a := cond_a AND input_valid_a;
IF NOT input_valid_a THEN
    channel_fault_a := channel_fault_a + 1;
END_IF;
cond_b := LimitHigh(raw_062_b, 122);
cond_b := cond_b AND quality_b;
cond_b := cond_b AND (NOT bypass_b);
input_valid_b := InputValid(raw_062_b, 0, 1000);
cond_b := cond_b AND input_valid_b;
IF NOT input_valid_b THEN
    channel_fault_b := channel_fault_b + 1;
END_IF;
cond_c := LimitHigh(raw_062_c, 122);
cond_c := cond_c AND quality_c;
cond_c := cond_c AND (NOT bypass_c);
input_valid_c := InputValid(raw_062_c, 0, 1000);
cond_c := cond_c AND input_valid_c;
IF NOT input_valid_c THEN
    channel_fault_c := channel_fault_c + 1;
END_IF;
cond_d := LimitHigh(raw_062_d, 122);
cond_d := cond_d AND quality_d;
cond_d := cond_d AND (NOT bypass_d);
input_valid_d := InputValid(raw_062_d, 0, 1000);
cond_d := cond_d AND input_valid_d;
IF NOT input_valid_d THEN
    channel_fault_d := channel_fault_d + 1;
END_IF;
vote_ok := TwoOfFour(cond_a, cond_b, cond_c, cond_d);
IF cond_a <> cond_b THEN
    diagnosis_count := diagnosis_count + 1;
END_IF;
IF cond_c <> cond_d THEN
    diagnosis_count := diagnosis_count + 1;
END_IF;
IF NOT vote_ok THEN
    diagnosis_count := diagnosis_count + 1;
END_IF;
latch_a_062 := RS_Next(vote_ok, train_a_reset, latch_a_062);
IF latch_a_062 AND (NOT train_a_inhibit) THEN
    mask_a_07 := mask_a_07 + 64;
    trip_a := 0 < 1;
    scram_a := 0 < 1;
    breaker_a := 0 > 1;
    mfw_a := 0 < 1;
    alarm_a := 0 < 1;
END_IF;
latch_b_062 := RS_Next(vote_ok, train_b_reset, latch_b_062);
IF latch_b_062 AND (NOT train_b_inhibit) THEN
    mask_b_07 := mask_b_07 + 64;
    trip_b := 0 < 1;
    scram_b := 0 < 1;
    breaker_b := 0 > 1;
    mfw_b := 0 < 1;
    alarm_b := 0 < 1;
END_IF;
IF (raw_062_a > 122) AND (NOT cond_a) THEN
    channel_fault_a := channel_fault_a + 1;
END_IF;
IF (raw_062_b > 122) AND (NOT cond_b) THEN
    channel_fault_b := channel_fault_b + 1;
END_IF;
IF (raw_062_c > 122) AND (NOT cond_c) THEN
    channel_fault_c := channel_fault_c + 1;
END_IF;
IF (raw_062_d > 122) AND (NOT cond_d) THEN
    channel_fault_d := channel_fault_d + 1;
END_IF;
IF vote_ok AND train_a_inhibit THEN
    diagnosis_count := diagnosis_count + 1;
END_IF;
IF vote_ok AND train_b_inhibit THEN
    diagnosis_count := diagnosis_count + 1;
END_IF;

cond_a := LimitHigh(raw_063_a, 123);
cond_a := cond_a AND quality_a;
cond_a := cond_a AND (NOT bypass_a);
input_valid_a := InputValid(raw_063_a, 0, 1000);
cond_a := cond_a AND input_valid_a;
IF NOT input_valid_a THEN
    channel_fault_a := channel_fault_a + 1;
END_IF;
cond_b := LimitHigh(raw_063_b, 123);
cond_b := cond_b AND quality_b;
cond_b := cond_b AND (NOT bypass_b);
input_valid_b := InputValid(raw_063_b, 0, 1000);
cond_b := cond_b AND input_valid_b;
IF NOT input_valid_b THEN
    channel_fault_b := channel_fault_b + 1;
END_IF;
cond_c := LimitHigh(raw_063_c, 123);
cond_c := cond_c AND quality_c;
cond_c := cond_c AND (NOT bypass_c);
input_valid_c := InputValid(raw_063_c, 0, 1000);
cond_c := cond_c AND input_valid_c;
IF NOT input_valid_c THEN
    channel_fault_c := channel_fault_c + 1;
END_IF;
cond_d := LimitHigh(raw_063_d, 123);
cond_d := cond_d AND quality_d;
cond_d := cond_d AND (NOT bypass_d);
input_valid_d := InputValid(raw_063_d, 0, 1000);
cond_d := cond_d AND input_valid_d;
IF NOT input_valid_d THEN
    channel_fault_d := channel_fault_d + 1;
END_IF;
vote_ok := TwoOfFour(cond_a, cond_b, cond_c, cond_d);
IF cond_a <> cond_b THEN
    diagnosis_count := diagnosis_count + 1;
END_IF;
IF cond_c <> cond_d THEN
    diagnosis_count := diagnosis_count + 1;
END_IF;
IF NOT vote_ok THEN
    diagnosis_count := diagnosis_count + 1;
END_IF;
latch_a_063 := RS_Next(vote_ok, train_a_reset, latch_a_063);
IF latch_a_063 AND (NOT train_a_inhibit) THEN
    mask_a_07 := mask_a_07 + 128;
    trip_a := 0 < 1;
    scram_a := 0 < 1;
    breaker_a := 0 > 1;
    afw_a := 0 < 1;
    alarm_a := 0 < 1;
END_IF;
latch_b_063 := RS_Next(vote_ok, train_b_reset, latch_b_063);
IF latch_b_063 AND (NOT train_b_inhibit) THEN
    mask_b_07 := mask_b_07 + 128;
    trip_b := 0 < 1;
    scram_b := 0 < 1;
    breaker_b := 0 > 1;
    afw_b := 0 < 1;
    alarm_b := 0 < 1;
END_IF;
IF (raw_063_a > 123) AND (NOT cond_a) THEN
    channel_fault_a := channel_fault_a + 1;
END_IF;
IF (raw_063_b > 123) AND (NOT cond_b) THEN
    channel_fault_b := channel_fault_b + 1;
END_IF;
IF (raw_063_c > 123) AND (NOT cond_c) THEN
    channel_fault_c := channel_fault_c + 1;
END_IF;
IF (raw_063_d > 123) AND (NOT cond_d) THEN
    channel_fault_d := channel_fault_d + 1;
END_IF;
IF vote_ok AND train_a_inhibit THEN
    diagnosis_count := diagnosis_count + 1;
END_IF;
IF vote_ok AND train_b_inhibit THEN
    diagnosis_count := diagnosis_count + 1;
END_IF;

cond_a := LimitHigh(raw_064_a, 124);
cond_a := cond_a AND quality_a;
cond_a := cond_a AND (NOT bypass_a);
input_valid_a := InputValid(raw_064_a, 0, 1000);
cond_a := cond_a AND input_valid_a;
IF NOT input_valid_a THEN
    channel_fault_a := channel_fault_a + 1;
END_IF;
cond_b := LimitHigh(raw_064_b, 124);
cond_b := cond_b AND quality_b;
cond_b := cond_b AND (NOT bypass_b);
input_valid_b := InputValid(raw_064_b, 0, 1000);
cond_b := cond_b AND input_valid_b;
IF NOT input_valid_b THEN
    channel_fault_b := channel_fault_b + 1;
END_IF;
cond_c := LimitHigh(raw_064_c, 124);
cond_c := cond_c AND quality_c;
cond_c := cond_c AND (NOT bypass_c);
input_valid_c := InputValid(raw_064_c, 0, 1000);
cond_c := cond_c AND input_valid_c;
IF NOT input_valid_c THEN
    channel_fault_c := channel_fault_c + 1;
END_IF;
cond_d := LimitHigh(raw_064_d, 124);
cond_d := cond_d AND quality_d;
cond_d := cond_d AND (NOT bypass_d);
input_valid_d := InputValid(raw_064_d, 0, 1000);
cond_d := cond_d AND input_valid_d;
IF NOT input_valid_d THEN
    channel_fault_d := channel_fault_d + 1;
END_IF;
vote_ok := TwoOfFour(cond_a, cond_b, cond_c, cond_d);
IF cond_a <> cond_b THEN
    diagnosis_count := diagnosis_count + 1;
END_IF;
IF cond_c <> cond_d THEN
    diagnosis_count := diagnosis_count + 1;
END_IF;
IF NOT vote_ok THEN
    diagnosis_count := diagnosis_count + 1;
END_IF;
latch_a_064 := RS_Next(vote_ok, train_a_reset, latch_a_064);
IF latch_a_064 AND (NOT train_a_inhibit) THEN
    mask_a_08 := mask_a_08 + 1;
    trip_a := 0 < 1;
    scram_a := 0 < 1;
    breaker_a := 0 > 1;
    si_a := 0 < 1;
    alarm_a := 0 < 1;
END_IF;
latch_b_064 := RS_Next(vote_ok, train_b_reset, latch_b_064);
IF latch_b_064 AND (NOT train_b_inhibit) THEN
    mask_b_08 := mask_b_08 + 1;
    trip_b := 0 < 1;
    scram_b := 0 < 1;
    breaker_b := 0 > 1;
    si_b := 0 < 1;
    alarm_b := 0 < 1;
END_IF;
IF (raw_064_a > 124) AND (NOT cond_a) THEN
    channel_fault_a := channel_fault_a + 1;
END_IF;
IF (raw_064_b > 124) AND (NOT cond_b) THEN
    channel_fault_b := channel_fault_b + 1;
END_IF;
IF (raw_064_c > 124) AND (NOT cond_c) THEN
    channel_fault_c := channel_fault_c + 1;
END_IF;
IF (raw_064_d > 124) AND (NOT cond_d) THEN
    channel_fault_d := channel_fault_d + 1;
END_IF;
IF vote_ok AND train_a_inhibit THEN
    diagnosis_count := diagnosis_count + 1;
END_IF;
IF vote_ok AND train_b_inhibit THEN
    diagnosis_count := diagnosis_count + 1;
END_IF;

cond_a := LimitHigh(raw_065_a, 125);
cond_a := cond_a AND quality_a;
cond_a := cond_a AND (NOT bypass_a);
input_valid_a := InputValid(raw_065_a, 0, 1000);
cond_a := cond_a AND input_valid_a;
IF NOT input_valid_a THEN
    channel_fault_a := channel_fault_a + 1;
END_IF;
cond_b := LimitHigh(raw_065_b, 125);
cond_b := cond_b AND quality_b;
cond_b := cond_b AND (NOT bypass_b);
input_valid_b := InputValid(raw_065_b, 0, 1000);
cond_b := cond_b AND input_valid_b;
IF NOT input_valid_b THEN
    channel_fault_b := channel_fault_b + 1;
END_IF;
cond_c := LimitHigh(raw_065_c, 125);
cond_c := cond_c AND quality_c;
cond_c := cond_c AND (NOT bypass_c);
input_valid_c := InputValid(raw_065_c, 0, 1000);
cond_c := cond_c AND input_valid_c;
IF NOT input_valid_c THEN
    channel_fault_c := channel_fault_c + 1;
END_IF;
cond_d := LimitHigh(raw_065_d, 125);
cond_d := cond_d AND quality_d;
cond_d := cond_d AND (NOT bypass_d);
input_valid_d := InputValid(raw_065_d, 0, 1000);
cond_d := cond_d AND input_valid_d;
IF NOT input_valid_d THEN
    channel_fault_d := channel_fault_d + 1;
END_IF;
vote_ok := TwoOfFour(cond_a, cond_b, cond_c, cond_d);
IF cond_a <> cond_b THEN
    diagnosis_count := diagnosis_count + 1;
END_IF;
IF cond_c <> cond_d THEN
    diagnosis_count := diagnosis_count + 1;
END_IF;
IF NOT vote_ok THEN
    diagnosis_count := diagnosis_count + 1;
END_IF;
latch_a_065 := RS_Next(vote_ok, train_a_reset, latch_a_065);
IF latch_a_065 AND (NOT train_a_inhibit) THEN
    mask_a_08 := mask_a_08 + 2;
    trip_a := 0 < 1;
    scram_a := 0 < 1;
    breaker_a := 0 > 1;
    ci_a := 0 < 1;
    alarm_a := 0 < 1;
END_IF;
latch_b_065 := RS_Next(vote_ok, train_b_reset, latch_b_065);
IF latch_b_065 AND (NOT train_b_inhibit) THEN
    mask_b_08 := mask_b_08 + 2;
    trip_b := 0 < 1;
    scram_b := 0 < 1;
    breaker_b := 0 > 1;
    ci_b := 0 < 1;
    alarm_b := 0 < 1;
END_IF;
IF (raw_065_a > 125) AND (NOT cond_a) THEN
    channel_fault_a := channel_fault_a + 1;
END_IF;
IF (raw_065_b > 125) AND (NOT cond_b) THEN
    channel_fault_b := channel_fault_b + 1;
END_IF;
IF (raw_065_c > 125) AND (NOT cond_c) THEN
    channel_fault_c := channel_fault_c + 1;
END_IF;
IF (raw_065_d > 125) AND (NOT cond_d) THEN
    channel_fault_d := channel_fault_d + 1;
END_IF;
IF vote_ok AND train_a_inhibit THEN
    diagnosis_count := diagnosis_count + 1;
END_IF;
IF vote_ok AND train_b_inhibit THEN
    diagnosis_count := diagnosis_count + 1;
END_IF;

cond_a := LimitHigh(raw_066_a, 126);
cond_a := cond_a AND quality_a;
cond_a := cond_a AND (NOT bypass_a);
input_valid_a := InputValid(raw_066_a, 0, 1000);
cond_a := cond_a AND input_valid_a;
IF NOT input_valid_a THEN
    channel_fault_a := channel_fault_a + 1;
END_IF;
cond_b := LimitHigh(raw_066_b, 126);
cond_b := cond_b AND quality_b;
cond_b := cond_b AND (NOT bypass_b);
input_valid_b := InputValid(raw_066_b, 0, 1000);
cond_b := cond_b AND input_valid_b;
IF NOT input_valid_b THEN
    channel_fault_b := channel_fault_b + 1;
END_IF;
cond_c := LimitHigh(raw_066_c, 126);
cond_c := cond_c AND quality_c;
cond_c := cond_c AND (NOT bypass_c);
input_valid_c := InputValid(raw_066_c, 0, 1000);
cond_c := cond_c AND input_valid_c;
IF NOT input_valid_c THEN
    channel_fault_c := channel_fault_c + 1;
END_IF;
cond_d := LimitHigh(raw_066_d, 126);
cond_d := cond_d AND quality_d;
cond_d := cond_d AND (NOT bypass_d);
input_valid_d := InputValid(raw_066_d, 0, 1000);
cond_d := cond_d AND input_valid_d;
IF NOT input_valid_d THEN
    channel_fault_d := channel_fault_d + 1;
END_IF;
vote_ok := TwoOfFour(cond_a, cond_b, cond_c, cond_d);
IF cond_a <> cond_b THEN
    diagnosis_count := diagnosis_count + 1;
END_IF;
IF cond_c <> cond_d THEN
    diagnosis_count := diagnosis_count + 1;
END_IF;
IF NOT vote_ok THEN
    diagnosis_count := diagnosis_count + 1;
END_IF;
latch_a_066 := RS_Next(vote_ok, train_a_reset, latch_a_066);
IF latch_a_066 AND (NOT train_a_inhibit) THEN
    mask_a_08 := mask_a_08 + 4;
    trip_a := 0 < 1;
    scram_a := 0 < 1;
    breaker_a := 0 > 1;
    mfw_a := 0 < 1;
    alarm_a := 0 < 1;
END_IF;
latch_b_066 := RS_Next(vote_ok, train_b_reset, latch_b_066);
IF latch_b_066 AND (NOT train_b_inhibit) THEN
    mask_b_08 := mask_b_08 + 4;
    trip_b := 0 < 1;
    scram_b := 0 < 1;
    breaker_b := 0 > 1;
    mfw_b := 0 < 1;
    alarm_b := 0 < 1;
END_IF;
IF (raw_066_a > 126) AND (NOT cond_a) THEN
    channel_fault_a := channel_fault_a + 1;
END_IF;
IF (raw_066_b > 126) AND (NOT cond_b) THEN
    channel_fault_b := channel_fault_b + 1;
END_IF;
IF (raw_066_c > 126) AND (NOT cond_c) THEN
    channel_fault_c := channel_fault_c + 1;
END_IF;
IF (raw_066_d > 126) AND (NOT cond_d) THEN
    channel_fault_d := channel_fault_d + 1;
END_IF;
IF vote_ok AND train_a_inhibit THEN
    diagnosis_count := diagnosis_count + 1;
END_IF;
IF vote_ok AND train_b_inhibit THEN
    diagnosis_count := diagnosis_count + 1;
END_IF;

cond_a := LimitHigh(raw_067_a, 127);
cond_a := cond_a AND quality_a;
cond_a := cond_a AND (NOT bypass_a);
input_valid_a := InputValid(raw_067_a, 0, 1000);
cond_a := cond_a AND input_valid_a;
IF NOT input_valid_a THEN
    channel_fault_a := channel_fault_a + 1;
END_IF;
cond_b := LimitHigh(raw_067_b, 127);
cond_b := cond_b AND quality_b;
cond_b := cond_b AND (NOT bypass_b);
input_valid_b := InputValid(raw_067_b, 0, 1000);
cond_b := cond_b AND input_valid_b;
IF NOT input_valid_b THEN
    channel_fault_b := channel_fault_b + 1;
END_IF;
cond_c := LimitHigh(raw_067_c, 127);
cond_c := cond_c AND quality_c;
cond_c := cond_c AND (NOT bypass_c);
input_valid_c := InputValid(raw_067_c, 0, 1000);
cond_c := cond_c AND input_valid_c;
IF NOT input_valid_c THEN
    channel_fault_c := channel_fault_c + 1;
END_IF;
cond_d := LimitHigh(raw_067_d, 127);
cond_d := cond_d AND quality_d;
cond_d := cond_d AND (NOT bypass_d);
input_valid_d := InputValid(raw_067_d, 0, 1000);
cond_d := cond_d AND input_valid_d;
IF NOT input_valid_d THEN
    channel_fault_d := channel_fault_d + 1;
END_IF;
vote_ok := TwoOfFour(cond_a, cond_b, cond_c, cond_d);
IF cond_a <> cond_b THEN
    diagnosis_count := diagnosis_count + 1;
END_IF;
IF cond_c <> cond_d THEN
    diagnosis_count := diagnosis_count + 1;
END_IF;
IF NOT vote_ok THEN
    diagnosis_count := diagnosis_count + 1;
END_IF;
latch_a_067 := RS_Next(vote_ok, train_a_reset, latch_a_067);
IF latch_a_067 AND (NOT train_a_inhibit) THEN
    mask_a_08 := mask_a_08 + 8;
    trip_a := 0 < 1;
    scram_a := 0 < 1;
    breaker_a := 0 > 1;
    afw_a := 0 < 1;
    alarm_a := 0 < 1;
END_IF;
latch_b_067 := RS_Next(vote_ok, train_b_reset, latch_b_067);
IF latch_b_067 AND (NOT train_b_inhibit) THEN
    mask_b_08 := mask_b_08 + 8;
    trip_b := 0 < 1;
    scram_b := 0 < 1;
    breaker_b := 0 > 1;
    afw_b := 0 < 1;
    alarm_b := 0 < 1;
END_IF;
IF (raw_067_a > 127) AND (NOT cond_a) THEN
    channel_fault_a := channel_fault_a + 1;
END_IF;
IF (raw_067_b > 127) AND (NOT cond_b) THEN
    channel_fault_b := channel_fault_b + 1;
END_IF;
IF (raw_067_c > 127) AND (NOT cond_c) THEN
    channel_fault_c := channel_fault_c + 1;
END_IF;
IF (raw_067_d > 127) AND (NOT cond_d) THEN
    channel_fault_d := channel_fault_d + 1;
END_IF;
IF vote_ok AND train_a_inhibit THEN
    diagnosis_count := diagnosis_count + 1;
END_IF;
IF vote_ok AND train_b_inhibit THEN
    diagnosis_count := diagnosis_count + 1;
END_IF;

cond_a := LimitHigh(raw_068_a, 128);
cond_a := cond_a AND quality_a;
cond_a := cond_a AND (NOT bypass_a);
input_valid_a := InputValid(raw_068_a, 0, 1000);
cond_a := cond_a AND input_valid_a;
IF NOT input_valid_a THEN
    channel_fault_a := channel_fault_a + 1;
END_IF;
cond_b := LimitHigh(raw_068_b, 128);
cond_b := cond_b AND quality_b;
cond_b := cond_b AND (NOT bypass_b);
input_valid_b := InputValid(raw_068_b, 0, 1000);
cond_b := cond_b AND input_valid_b;
IF NOT input_valid_b THEN
    channel_fault_b := channel_fault_b + 1;
END_IF;
cond_c := LimitHigh(raw_068_c, 128);
cond_c := cond_c AND quality_c;
cond_c := cond_c AND (NOT bypass_c);
input_valid_c := InputValid(raw_068_c, 0, 1000);
cond_c := cond_c AND input_valid_c;
IF NOT input_valid_c THEN
    channel_fault_c := channel_fault_c + 1;
END_IF;
cond_d := LimitHigh(raw_068_d, 128);
cond_d := cond_d AND quality_d;
cond_d := cond_d AND (NOT bypass_d);
input_valid_d := InputValid(raw_068_d, 0, 1000);
cond_d := cond_d AND input_valid_d;
IF NOT input_valid_d THEN
    channel_fault_d := channel_fault_d + 1;
END_IF;
vote_ok := TwoOfFour(cond_a, cond_b, cond_c, cond_d);
IF cond_a <> cond_b THEN
    diagnosis_count := diagnosis_count + 1;
END_IF;
IF cond_c <> cond_d THEN
    diagnosis_count := diagnosis_count + 1;
END_IF;
IF NOT vote_ok THEN
    diagnosis_count := diagnosis_count + 1;
END_IF;
latch_a_068 := RS_Next(vote_ok, train_a_reset, latch_a_068);
IF latch_a_068 AND (NOT train_a_inhibit) THEN
    mask_a_08 := mask_a_08 + 16;
    trip_a := 0 < 1;
    scram_a := 0 < 1;
    breaker_a := 0 > 1;
    si_a := 0 < 1;
    alarm_a := 0 < 1;
END_IF;
latch_b_068 := RS_Next(vote_ok, train_b_reset, latch_b_068);
IF latch_b_068 AND (NOT train_b_inhibit) THEN
    mask_b_08 := mask_b_08 + 16;
    trip_b := 0 < 1;
    scram_b := 0 < 1;
    breaker_b := 0 > 1;
    si_b := 0 < 1;
    alarm_b := 0 < 1;
END_IF;
IF (raw_068_a > 128) AND (NOT cond_a) THEN
    channel_fault_a := channel_fault_a + 1;
END_IF;
IF (raw_068_b > 128) AND (NOT cond_b) THEN
    channel_fault_b := channel_fault_b + 1;
END_IF;
IF (raw_068_c > 128) AND (NOT cond_c) THEN
    channel_fault_c := channel_fault_c + 1;
END_IF;
IF (raw_068_d > 128) AND (NOT cond_d) THEN
    channel_fault_d := channel_fault_d + 1;
END_IF;
IF vote_ok AND train_a_inhibit THEN
    diagnosis_count := diagnosis_count + 1;
END_IF;
IF vote_ok AND train_b_inhibit THEN
    diagnosis_count := diagnosis_count + 1;
END_IF;

cond_a := LimitHigh(raw_069_a, 129);
cond_a := cond_a AND quality_a;
cond_a := cond_a AND (NOT bypass_a);
input_valid_a := InputValid(raw_069_a, 0, 1000);
cond_a := cond_a AND input_valid_a;
IF NOT input_valid_a THEN
    channel_fault_a := channel_fault_a + 1;
END_IF;
cond_b := LimitHigh(raw_069_b, 129);
cond_b := cond_b AND quality_b;
cond_b := cond_b AND (NOT bypass_b);
input_valid_b := InputValid(raw_069_b, 0, 1000);
cond_b := cond_b AND input_valid_b;
IF NOT input_valid_b THEN
    channel_fault_b := channel_fault_b + 1;
END_IF;
cond_c := LimitHigh(raw_069_c, 129);
cond_c := cond_c AND quality_c;
cond_c := cond_c AND (NOT bypass_c);
input_valid_c := InputValid(raw_069_c, 0, 1000);
cond_c := cond_c AND input_valid_c;
IF NOT input_valid_c THEN
    channel_fault_c := channel_fault_c + 1;
END_IF;
cond_d := LimitHigh(raw_069_d, 129);
cond_d := cond_d AND quality_d;
cond_d := cond_d AND (NOT bypass_d);
input_valid_d := InputValid(raw_069_d, 0, 1000);
cond_d := cond_d AND input_valid_d;
IF NOT input_valid_d THEN
    channel_fault_d := channel_fault_d + 1;
END_IF;
vote_ok := TwoOfFour(cond_a, cond_b, cond_c, cond_d);
IF cond_a <> cond_b THEN
    diagnosis_count := diagnosis_count + 1;
END_IF;
IF cond_c <> cond_d THEN
    diagnosis_count := diagnosis_count + 1;
END_IF;
IF NOT vote_ok THEN
    diagnosis_count := diagnosis_count + 1;
END_IF;
latch_a_069 := RS_Next(vote_ok, train_a_reset, latch_a_069);
IF latch_a_069 AND (NOT train_a_inhibit) THEN
    mask_a_08 := mask_a_08 + 32;
    trip_a := 0 < 1;
    scram_a := 0 < 1;
    breaker_a := 0 > 1;
    ci_a := 0 < 1;
    alarm_a := 0 < 1;
END_IF;
latch_b_069 := RS_Next(vote_ok, train_b_reset, latch_b_069);
IF latch_b_069 AND (NOT train_b_inhibit) THEN
    mask_b_08 := mask_b_08 + 32;
    trip_b := 0 < 1;
    scram_b := 0 < 1;
    breaker_b := 0 > 1;
    ci_b := 0 < 1;
    alarm_b := 0 < 1;
END_IF;
IF (raw_069_a > 129) AND (NOT cond_a) THEN
    channel_fault_a := channel_fault_a + 1;
END_IF;
IF (raw_069_b > 129) AND (NOT cond_b) THEN
    channel_fault_b := channel_fault_b + 1;
END_IF;
IF (raw_069_c > 129) AND (NOT cond_c) THEN
    channel_fault_c := channel_fault_c + 1;
END_IF;
IF (raw_069_d > 129) AND (NOT cond_d) THEN
    channel_fault_d := channel_fault_d + 1;
END_IF;
IF vote_ok AND train_a_inhibit THEN
    diagnosis_count := diagnosis_count + 1;
END_IF;
IF vote_ok AND train_b_inhibit THEN
    diagnosis_count := diagnosis_count + 1;
END_IF;
